// TIA Portal project "智能配药稳定版" (V16)

(* hardware
DEVICE "S7-1200 station_1"  S7-1200 Station
   slot 0: "Rack_0"  S7-1200 Rack  Rack  V1.0
   slot 1: "1.自动供料单元"  CPU 1214C DC/DC/DC  6ES7 214-1AG40-0XB0  V4.4
DEVICE "GSD device_1"  GSD.Device.PN
   slot 0: "机架"  Rack  V1.0
   slot 0: "DEC"  EX-1110  02-01-05  V10.00.00
      slot 0: "TPS Development Toolkit Drivertest"  TPS Development Toolkit Drivertest
      slot 1: "PN-IO"  PN-IO
         slot 1: "Port 1 - RJ45"  Port 1 - RJ45
         slot 2: "Port 2 - RJ45"  Port 2 - RJ45
   slot 1: "EX_210H_1"  EX_210H  1.0
      slot 0: "EX_210H"  EX_210H
   slot 2: "EX_2108_1"  EX_2108  1.0
      slot 0: "EX_2108"  EX_2108
   slot 3: "EX_3208_1"  EX_3208  1.0
      slot 0: "EX_3208"  EX_3208
DEVICE "1.自动供料单元_HMI"  KTP700 Basic PN
   slot 0: "2.自动供料单元_HMI"  KTP700 Basic PN  6AV2 123-2GB03-0AX0  16.0.0.0
   slot 1: "HMI_RT_1"  KTP700 Basic PN  6AV2 123-2GB03-0AX0  16.0.0.0
   slot 5: "2.自动供料单元_HMI.IE_CP_1"  PROFINET Interface  16.0.0.0
      slot 1: "PROFINET Interface_1"  PROFINET Interface
         slot 1: "Port_1"  Port
DEVICE "GSD device_2"  GSD.Device.PN
   slot 0: "机架"  Rack  V1.0
   slot 0: "SINAMICS-V90-PN"  SINAMICS V90 PN V1.0  6SL3 210-5Fxxx-xxFx  V1.00
      slot 0: "SINAMICS V90 PN V1.0"  SINAMICS V90 PN V1.0
      slot 1: "PN-IO"  PN-IO
         slot 1: "端口1"  Port 1
         slot 2: "端口2"  Port 2
      slot 1: "驱动_1"  DRIVE OBJECT
         slot 0: "模块访问点"  Module Access Point
         slot 1: "没有 PROFIsafe"  without PROFIsafe
   slot 2: "标准报文3, PZD-5/9"  Standard telegram 3, PZD 5/9
DEVICE "S7-1200 station_2"  S7-1200 Station
   slot 0: "Rack_0"  S7-1200 Rack  Rack  V1.0
   slot 1: "2.智能分拣单元"  CPU 1214C DC/DC/DC  6ES7 214-1AG40-0XB0  V4.4
DEVICE "2.智能分拣单元_HMI"  KTP700 Basic PN
   slot 0: "HMI_1"  KTP700 Basic PN  6AV2 123-2GB03-0AX0  16.0.0.0
   slot 1: "HMI_RT_2"  KTP700 Basic PN  6AV2 123-2GB03-0AX0  16.0.0.0
   slot 5: "HMI_1.IE_CP_1"  PROFINET Interface  16.0.0.0
      slot 1: "PROFINET Interface_1"  PROFINET Interface
         slot 1: "Port_1"  Port
DEVICE "S7-1200 station_3"  S7-1200 Station
   slot 0: "Rack_0"  S7-1200 Rack  Rack  V1.0
   slot 1: "3.智能仓储单元"  CPU 1214C DC/DC/DC  6ES7 214-1AG40-0XB0  V4.4
   slot 2: "SM 1278_1"  4SI IO link  6ES7 278-4BD32-0XB0  V2.1
   slot 3: "CB 1241 (RS485)"  CB 1241 (RS485)  6ES7 241-1CH30-1XB0  V1.0
   slot 101: "CM 1243-5"  CM 1243-5  6GK7 243-5DX30-0XE0  V1.3
DEVICE "3.智能仓储单元_HMI"  KTP700 Basic PN
   slot 0: "3.智能仓储单元_HMI"  KTP700 Basic PN  6AV2 123-2GB03-0AX0  16.0.0.0
   slot 1: "HMI_RT_3"  KTP700 Basic PN  6AV2 123-2GB03-0AX0  16.0.0.0
   slot 5: "3.智能仓储单元_HMI.IE_CP_1"  PROFINET Interface  16.0.0.0
      slot 1: "PROFINET Interface_1"  PROFINET Interface
         slot 1: "Port_1"  Port
DEVICE "GSD device_3"  GSD.Device.PN
   slot 0: "机架"  Rack  V1.0
   slot 0: "DEC_1"  EX-1110  02-01-05  V10.00.00
      slot 0: "TPS Development Toolkit Drivertest"  TPS Development Toolkit Drivertest
      slot 1: "PN-IO"  PN-IO
         slot 1: "Port 1 - RJ45"  Port 1 - RJ45
         slot 2: "Port 2 - RJ45"  Port 2 - RJ45
   slot 1: "EX_210H_1"  EX_210H  1.0
      slot 0: "EX_210H"  EX_210H
   slot 2: "EX_3208_1"  EX_3208  1.0
      slot 0: "EX_3208"  EX_3208
DEVICE "GSD device_4"  GSD.Device.PN
   slot 0: "机架"  Rack  V1.0
   slot 0: "SINAMICS-V90-PN_1"  SINAMICS V90 PN V1.0  6SL3 210-5Fxxx-xxFx  V1.00
      slot 0: "SINAMICS V90 PN V1.0"  SINAMICS V90 PN V1.0
      slot 1: "PN-IO"  PN-IO
         slot 1: "端口1"  Port 1
         slot 2: "端口2"  Port 2
      slot 1: "驱动_1"  DRIVE OBJECT
         slot 0: "模块访问点"  Module Access Point
         slot 1: "没有 PROFIsafe"  without PROFIsafe
   slot 2: "标准报文3, PZD-5/9"  Standard telegram 3, PZD 5/9
DEVICE "GSD device_5"  GSD.Device.PN
   slot 0: "机架"  Rack  V1.0
   slot 0: "SINAMICS-V90-PN_2"  SINAMICS V90 PN V1.0  6SL3 210-5Fxxx-xxFx  V1.00
      slot 0: "SINAMICS V90 PN V1.0"  SINAMICS V90 PN V1.0
      slot 1: "PN-IO"  PN-IO
         slot 1: "端口1"  Port 1
         slot 2: "端口2"  Port 2
      slot 1: "驱动_1"  DRIVE OBJECT
         slot 0: "模块访问点"  Module Access Point
         slot 1: "没有 PROFIsafe"  without PROFIsafe
   slot 2: "标准报文3, PZD-5/9"  Standard telegram 3, PZD 5/9
DEVICE "GSD device_6"  GSD.Device
   slot 0: "机架_0"  Rail
   slot 0: "Slave_1"  DP-Slave_1  Z1.0
DEVICE "GSD device_7"  GSD.Device.PN
   slot 0: "机架"  Rack  V1.0
   slot 0: "DEC_2"  EX-1110  02-01-05  V10.00.00
      slot 0: "TPS Development Toolkit Drivertest"  TPS Development Toolkit Drivertest
      slot 1: "PN-IO"  PN-IO
         slot 1: "Port 1 - RJ45"  Port 1 - RJ45
         slot 2: "Port 2 - RJ45"  Port 2 - RJ45
   slot 1: "EX_210H_1"  EX_210H  1.0
      slot 0: "EX_210H"  EX_210H
   slot 2: "EX_210H_2"  EX_210H  1.0
      slot 0: "EX_210H"  EX_210H
   slot 3: "EX_3208_1"  EX_3208  1.0
      slot 0: "EX_3208"  EX_3208
   slot 4: "EX_3208_2"  EX_3208  1.0
      slot 0: "EX_3208"  EX_3208
DEVICE "S71500/ET200MP station_1"  S7-1500 station
   slot 0: "导轨_0"  Rack  6ES7 590-1***0-0AA0
   slot 1: "0.数据管理单元"  CPU 1511-1 PN  6ES7 511-1AK02-0AB0  V2.8
      slot 3: "CPU 显示_1"  6ES7591-1AA00-0AA0
      slot 32768: "PROFINET 接口_1"  X1
         slot 32769: "端口_1"  X1 P1
         slot 32770: "端口_2"  X1 P2
      slot 34817: "Virtual CP interface port_1"  Virtual CP interface port  Virtual CP interface port
   slot 2: "DI 16x24VDC / DQ 16x24VDC/0.5A BA_1"  DI 16x24VDC/DQ 16x24VDC/0.5A BA  6ES7 523-1BL00-0AA0  V1.1
DEVICE "GSD device_8"  GSD.Device.PN
   slot 0: "机架"  Rack  V1.0
   slot 0: "SG-GATEWAY"  Master(h750)  SG-PNMB-MS2.0  SW2.0.0
      slot 0: "Master(h750)"  Master(h750)
      slot 1: "X1"  X1
         slot 1: "X1 P1"  X1 P1
         slot 2: "X1 P2"  X1 P2
      slot 1: "Control and Status_1"  Control and Status
         slot 0: "Control and Status"  Control and Status
   slot 2: "03H Read 17 Regs_1"  03H Read 17 Regs
      slot 0: "03H Read 17 Regs"  03H Read 17 Regs
   slot 3: "03H Read 2 Regs_1"  03H Read 2 Regs
      slot 0: "03H Read 2 Regs"  03H Read 2 Regs
   slot 4: "10H Write 1 Reg_1"  10H Write 1 Reg
      slot 0: "10H Write 1 Reg"  10H Write 1 Reg
   slot 5: "03H Read 2 Regs_2"  03H Read 2 Regs
      slot 0: "03H Read 2 Regs"  03H Read 2 Regs
   slot 6: "05H ForceSingleCoil_1"  05H ForceSingleCoil
      slot 0: "05H ForceSingleCoil"  05H ForceSingleCoil
   slot 7: "05H ForceSingleCoil_2"  05H ForceSingleCoil
      slot 0: "05H ForceSingleCoil"  05H ForceSingleCoil
   slot 8: "05H ForceSingleCoil_3"  05H ForceSingleCoil
      slot 0: "05H ForceSingleCoil"  05H ForceSingleCoil
   slot 9: "05H ForceSingleCoil_4"  05H ForceSingleCoil
      slot 0: "05H ForceSingleCoil"  05H ForceSingleCoil
DEVICE "0.数据管理单元_HMI"  KTP700 Basic PN
   slot 0: "0.数据管理单元_HMI"  KTP700 Basic PN  6AV2 123-2GB03-0AX0  16.0.0.0
   slot 1: "HMI_RT_4"  KTP700 Basic PN  6AV2 123-2GB03-0AX0  16.0.0.0
   slot 5: "0.数据管理单元_HMI.IE_CP_1"  PROFINET Interface  16.0.0.0
      slot 1: "PROFINET Interface_1"  PROFINET Interface
         slot 1: "Port_1"  Port
*)

// ===== PLC "1.自动供料单元"  CPU 1214C DC/DC/DC =====

VAR_GLOBAL   // PLC tag table "默认变量表"
   "System_Byte" AT %MB501 : Byte;
   "FirstScan" AT %M501.0 : Bool;
   "DiagStatusUpdate" AT %M501.1 : Bool;
   "AlwaysTRUE" AT %M501.2 : Bool;
   "AlwaysFALSE" AT %M501.3 : Bool;
   "Clock_Byte" AT %MB500 : Byte;
   "Clock_10Hz" AT %M500.0 : Bool;
   "Clock_5Hz" AT %M500.1 : Bool;
   "Clock_2.5Hz" AT %M500.2 : Bool;
   "Clock_2Hz" AT %M500.3 : Bool;
   "Clock_1.25Hz" AT %M500.4 : Bool;
   "Clock_1Hz" AT %M500.5 : Bool;
   "Clock_0.625Hz" AT %M500.6 : Bool;
   "Clock_0.5Hz" AT %M500.7 : Bool;
   "数量检测沿1" AT %M10.0 : Bool;
   "数量检测沿2" AT %M10.1 : Bool;
   "数量检测沿3" AT %M10.2 : Bool;
   "Tag_1" AT %M11.0 : Bool;
   "Tag_2" AT %M11.1 : Bool;
   "Tag_3" AT %M11.2 : Bool;
END_VAR

VAR_GLOBAL   // PLC tag table "第一站变量表"
   "[100]伺服左极限" AT %I0.0 : Bool;
   "[101]伺服右极限" AT %I0.1 : Bool;
   "[102]伺服原点" AT %I0.2 : Bool;
   "[103]步进原点" AT %I0.3 : Bool;
   "[104]步进右极限" AT %I0.4 : Bool;
   "[105]启动" AT %I0.5 : Bool;
   "[106]停止" AT %I0.6 : Bool;
   "[107]复位" AT %I0.7 : Bool;
   "[110]急停" AT %I1.0 : Bool;
   "[111]手自动" AT %I1.1 : Bool;
   "[112]料仓有无料盒" AT %I1.2 : Bool;
   "[113]取料位有无料盒" AT %I1.3 : Bool;
   "[114]功能1" AT %I1.4 : Bool;
   "[115]功能2" AT %I1.5 : Bool;
   "[120]A库物料检测" AT %I2.0 : Bool;
   "[121]B库物料检测" AT %I2.1 : Bool;
   "[122]取料位有无料块" AT %I2.2 : Bool;
   "[123]转盘装配到位检测" AT %I2.3 : Bool;
   "[124]推料盒缩回位" AT %I2.4 : Bool;
   "[125]推料盒伸出位" AT %I2.5 : Bool;
   "[126]A推料伸出位" AT %I2.6 : Bool;
   "[127]A推料缩回位" AT %I2.7 : Bool;
   "[130]B推料伸出位" AT %I3.0 : Bool;
   "[131]B推料缩回位" AT %I3.1 : Bool;
   "[132]取料盒下降位" AT %I3.2 : Bool;
   "[133]取料盒上升位" AT %I3.3 : Bool;
   "[134]取料块伸出位" AT %I3.4 : Bool;
   "[135]取料块缩回位" AT %I3.5 : Bool;
   "[136]取料块下降位" AT %I3.6 : Bool;
   "[137]取料块上升位" AT %I3.7 : Bool;
   "[140]检测伸出位" AT %I4.0 : Bool;
   "[141]检测缩回位" AT %I4.1 : Bool;
   "[142]检测下降位" AT %I4.2 : Bool;
   "[143]检测上升位" AT %I4.3 : Bool;
   "[156]安全光栅" AT %I5.6 : Bool;
   "[164]深度检测当前值" AT %IW64 : Int;
   "轴_1_Drive_IN" AT %I68.0 : "PD_TEL3_IN";
   "[300]转盘步进脉冲" AT %Q0.0 : Bool;
   "[301]转盘步进方向" AT %Q0.1 : Bool;
   "[302]黄色指示灯" AT %Q0.2 : Bool;
   "[303]绿色指示灯" AT %Q0.3 : Bool;
   "[304]红色指示灯" AT %Q0.4 : Bool;
   "[305]转盘皮带电机(正转)" AT %Q0.5 : Bool;
   "[306]转盘皮带电机(反转)" AT %Q0.6 : Bool;
   "[307]声光报警" AT %Q0.7 : Bool;
   "[310]检测伸缩气缸" AT %Q1.0 : Bool;
   "[311]检测升降气缸" AT %Q1.1 : Bool;
   "[320]底盒推料气缸" AT %Q2.0 : Bool;
   "[322]B库推料气缸" AT %Q2.2 : Bool;
   "[323]取底盒升降气缸" AT %Q2.3 : Bool;
   "[324]取料块升降气缸" AT %Q2.4 : Bool;
   "[325]取料块伸缩气缸" AT %Q2.5 : Bool;
   "[326]取料盒夹爪" AT %Q2.6 : Bool;
   "[327]取料块吸盘" AT %Q2.7 : Bool;
   "轴_1_Drive_OUT" AT %Q64.0 : "PD_TEL3_OUT";
   "[144]机械手夹紧到位" AT %I4.4 : Bool;
   "[145]机械手松开到位" AT %I4.5 : Bool;
   "[321]A库推料气缸" AT %Q2.1 : Bool;
END_VAR

DATA_BLOCK "状态控制数据"   // DB33
{ S7_Optimized_Access := 'FALSE' }
VERSION : 0.1
   VAR
      在线状态 : Bool;   // PLC已经上电
      忙碌状态 : Bool;   // 一站已经接单
      空闲状态 : Bool;   // 一站准备就绪(没急停，初始化已经完成，光栅没被挡)
      故障状态 : Bool;   // 报警、光栅被挡
   END_VAR
BEGIN
END_DATA_BLOCK

DATA_BLOCK "初始化数据"   // DB34
{ S7_Optimized_Access := 'FALSE' }
VERSION : 0.1
   VAR
      手动模式 : Bool;
      自动模式 : Bool;
      自动运行模式 : Bool;
      急停状态 : Bool;
      安全光栅被挡 : Bool;
      红灯_内部 : Bool;
      黄灯_内部 : Bool;
      绿灯_内部 : Bool;
      初始化步骤 : Int;
      初始化条件 : Bool;
      初始化下降沿 : Bool;
      初始化中 : Bool;
      初始化故障 : Bool;
      初始化完成 : Bool;
      报警等级 : Int;
      报警确认按钮 : Bool;
      气缸报警复位 : Bool;
      底盒推料气缸报警 : Bool;
      A库推料气缸报警 : Bool;
      B库推料气缸报警 : Bool;
      检测伸缩气缸报警 : Bool;
      检测升降气缸报警 : Bool;
      取料块升降气缸报警 : Bool;
      取料块伸缩气缸报警 : Bool;
      取料盒夹爪报警 : Bool;
      气缸报警输出 : Bool;
      轴回零错误 : Bool;
      报警总输出 : Bool;
   END_VAR
BEGIN
END_DATA_BLOCK

// folder: System blocks/Program resources

DATA_BLOCK "吸住料块上升计时"   // DB10
{ S7_Optimized_Access := 'TRUE' }
AUTHOR : Simatic
FAMILY : IEC
NAME : IEC_TMR
VERSION : 1.0
// stored: InstanceOfName IEC_TIMER
"IEC_TIMER"
BEGIN
END_DATA_BLOCK

DATA_BLOCK "IEC_Timer_0_DB_10"   // DB14
{ S7_Optimized_Access := 'TRUE' }
AUTHOR : Simatic
FAMILY : IEC
NAME : IEC_TMR
VERSION : 1.0
// stored: InstanceOfName IEC_TIMER
"IEC_TIMER"
BEGIN
END_DATA_BLOCK

DATA_BLOCK "IEC_Timer_0_DB_5"   // DB16
{ S7_Optimized_Access := 'TRUE' }
AUTHOR : Simatic
FAMILY : IEC
NAME : IEC_TMR
VERSION : 1.0
// stored: InstanceOfName IEC_TIMER
"IEC_TIMER"
BEGIN
END_DATA_BLOCK

DATA_BLOCK "IEC_Timer_0_DB_2"   // DB19
{ S7_Optimized_Access := 'TRUE' }
AUTHOR : Simatic
FAMILY : IEC
NAME : IEC_TMR
VERSION : 1.0
// stored: InstanceOfName IEC_TIMER
"IEC_TIMER"
BEGIN
END_DATA_BLOCK

DATA_BLOCK "IEC_Timer_0_DB_3"   // DB21
{ S7_Optimized_Access := 'TRUE' }
AUTHOR : Simatic
FAMILY : IEC
NAME : IEC_TMR
VERSION : 1.0
// stored: InstanceOfName IEC_TIMER
"IEC_TIMER"
BEGIN
END_DATA_BLOCK

DATA_BLOCK "IEC_Timer_0_DB_7"   // DB23
{ S7_Optimized_Access := 'TRUE' }
AUTHOR : Simatic
FAMILY : IEC
NAME : IEC_TMR
VERSION : 1.0
// stored: InstanceOfName IEC_TIMER
"IEC_TIMER"
BEGIN
END_DATA_BLOCK

DATA_BLOCK "IEC_Timer_0_DB_6"   // DB24
{ S7_Optimized_Access := 'TRUE' }
AUTHOR : Simatic
FAMILY : IEC
NAME : IEC_TMR
VERSION : 1.0
// stored: InstanceOfName IEC_TIMER
"IEC_TIMER"
BEGIN
END_DATA_BLOCK

DATA_BLOCK "IEC_Timer_0_DB_8"   // DB25
{ S7_Optimized_Access := 'TRUE' }
AUTHOR : Simatic
FAMILY : IEC
NAME : IEC_TMR
VERSION : 1.0
// stored: InstanceOfName IEC_TIMER
"IEC_TIMER"
BEGIN
END_DATA_BLOCK

DATA_BLOCK "IEC_Timer_0_DB_9"   // DB26
{ S7_Optimized_Access := 'TRUE' }
AUTHOR : Simatic
FAMILY : IEC
NAME : IEC_TMR
VERSION : 1.0
// stored: InstanceOfName IEC_TIMER
"IEC_TIMER"
BEGIN
END_DATA_BLOCK

DATA_BLOCK "IEC_Timer_0_DB_11"   // DB27
{ S7_Optimized_Access := 'TRUE' }
AUTHOR : Simatic
FAMILY : IEC
NAME : IEC_TMR
VERSION : 1.0
// stored: InstanceOfName IEC_TIMER
"IEC_TIMER"
BEGIN
END_DATA_BLOCK

DATA_BLOCK "IEC_Timer_0_DB_12"   // DB28
{ S7_Optimized_Access := 'TRUE' }
AUTHOR : Simatic
FAMILY : IEC
NAME : IEC_TMR
VERSION : 1.0
// stored: InstanceOfName IEC_TIMER
"IEC_TIMER"
BEGIN
END_DATA_BLOCK

DATA_BLOCK "IEC_Timer_0_DB_13"   // DB29
{ S7_Optimized_Access := 'TRUE' }
AUTHOR : Simatic
FAMILY : IEC
NAME : IEC_TMR
VERSION : 1.0
// stored: InstanceOfName IEC_TIMER
"IEC_TIMER"
BEGIN
END_DATA_BLOCK

DATA_BLOCK "IEC_Timer_0_DB_14"   // DB30
{ S7_Optimized_Access := 'TRUE' }
AUTHOR : Simatic
FAMILY : IEC
NAME : IEC_TMR
VERSION : 1.0
// stored: InstanceOfName IEC_TIMER
"IEC_TIMER"
BEGIN
END_DATA_BLOCK

DATA_BLOCK "IEC_Timer_0_DB_15"   // DB31
{ S7_Optimized_Access := 'TRUE' }
AUTHOR : Simatic
FAMILY : IEC
NAME : IEC_TMR
VERSION : 1.0
// stored: InstanceOfName IEC_TIMER
"IEC_TIMER"
BEGIN
END_DATA_BLOCK

DATA_BLOCK "IEC_Timer_0_DB_4"   // DB32
{ S7_Optimized_Access := 'TRUE' }
AUTHOR : Simatic
FAMILY : IEC
NAME : IEC_TMR
VERSION : 1.0
// stored: InstanceOfName IEC_TIMER
"IEC_TIMER"
BEGIN
END_DATA_BLOCK

DATA_BLOCK "IEC_Timer_0_DB_23"   // DB35
{ S7_Optimized_Access := 'TRUE' }
AUTHOR : Simatic
FAMILY : IEC
NAME : IEC_TMR
VERSION : 1.0
// stored: InstanceOfName IEC_TIMER
"IEC_TIMER"
BEGIN
END_DATA_BLOCK

DATA_BLOCK "_1.自动供料单元_Receive_DB"   // DB38
{ S7_Optimized_Access := 'TRUE' }
AUTHOR : SIMATIC
FAMILY : MC7Plus
NAME : TC_IP_v4
VERSION : 1.0
// stored: InstanceOfName TCON_IP_v4
"TCON_IP_v4"
BEGIN
   ID := 105;
   InterfaceId := 64;
   LocalPort := 8899;
   RemotePort := 8899;
   RemoteAddress.ADDR[1] := 192;
   RemoteAddress.ADDR[2] := 168;
   RemoteAddress.ADDR[3] := 40;
   RemoteAddress.ADDR[4] := 100;
END_DATA_BLOCK

DATA_BLOCK "IEC_Timer_0_DB_24"   // DB39
{ S7_Optimized_Access := 'TRUE' }
AUTHOR : Simatic
FAMILY : IEC
NAME : IEC_TMR
VERSION : 1.0
// stored: InstanceOfName IEC_TIMER
"IEC_TIMER"
BEGIN
END_DATA_BLOCK

DATA_BLOCK "IEC_Timer_0_DB_16"   // DB40
{ S7_Optimized_Access := 'TRUE' }
AUTHOR : Simatic
FAMILY : IEC
NAME : IEC_TMR
VERSION : 1.0
// stored: InstanceOfName IEC_TIMER
"IEC_TIMER"
BEGIN
END_DATA_BLOCK

DATA_BLOCK "IEC_Timer_0_DB_17"   // DB41
{ S7_Optimized_Access := 'TRUE' }
AUTHOR : Simatic
FAMILY : IEC
NAME : IEC_TMR
VERSION : 1.0
// stored: InstanceOfName IEC_TIMER
"IEC_TIMER"
BEGIN
END_DATA_BLOCK

DATA_BLOCK "IEC_Timer_0_DB_18"   // DB42
{ S7_Optimized_Access := 'TRUE' }
AUTHOR : Simatic
FAMILY : IEC
NAME : IEC_TMR
VERSION : 1.0
// stored: InstanceOfName IEC_TIMER
"IEC_TIMER"
BEGIN
END_DATA_BLOCK

DATA_BLOCK "IEC_Timer_0_DB_19"   // DB43
{ S7_Optimized_Access := 'TRUE' }
AUTHOR : Simatic
FAMILY : IEC
NAME : IEC_TMR
VERSION : 1.0
// stored: InstanceOfName IEC_TIMER
"IEC_TIMER"
BEGIN
END_DATA_BLOCK

DATA_BLOCK "IEC_Timer_0_DB_20"   // DB44
{ S7_Optimized_Access := 'TRUE' }
AUTHOR : Simatic
FAMILY : IEC
NAME : IEC_TMR
VERSION : 1.0
// stored: InstanceOfName IEC_TIMER
"IEC_TIMER"
BEGIN
END_DATA_BLOCK

DATA_BLOCK "IEC_Timer_0_DB_21"   // DB45
{ S7_Optimized_Access := 'TRUE' }
AUTHOR : Simatic
FAMILY : IEC
NAME : IEC_TMR
VERSION : 1.0
// stored: InstanceOfName IEC_TIMER
"IEC_TIMER"
BEGIN
END_DATA_BLOCK

DATA_BLOCK "IEC_Timer_0_DB_22"   // DB46
{ S7_Optimized_Access := 'TRUE' }
AUTHOR : Simatic
FAMILY : IEC
NAME : IEC_TMR
VERSION : 1.0
// stored: InstanceOfName IEC_TIMER
"IEC_TIMER"
BEGIN
END_DATA_BLOCK

// folder: 手动模式

DATA_BLOCK "手动模式数据"   // DB12
{ S7_Optimized_Access := 'FALSE' }
VERSION : 0.1
   VAR
      S10推料盒步骤 : Real;
      S20推料块步骤 : Real;
      S30放料块步骤 : Real;
      S40送料盒步骤 : Real;
      手动总步骤 : Real;
      料块仓选择 : Int := 1;
      沿1 : Bool;
      沿2 : Bool;
      沿3 : Bool;
      沿4 : Bool;
   END_VAR
BEGIN
END_DATA_BLOCK

// folder: 自动模式

DATA_BLOCK "自动模式数据"   // DB22
{ S7_Optimized_Access := 'FALSE' }
VERSION : 0.1
   VAR
      Z10步骤 : Real;
      Z20步骤 : Real;
      Z30步骤 : Real;
      Z40步骤 : Real;
      Z50步骤 : Real;
      自动模式总步骤 : Real;
      推料盒数 : Bool;
      开始信号 : Bool;
      ab物料选择 : Int;
      料盒使用数 : Int;
      a料使用数 : Int;
      b料使用数 : Int;
      当前深度检测_1 : Real;   // 模数转换
      当前深度检测_2 : Real;   // 模数转换
      当前深度检测 : Real;
      深度保存 : Array[0..1] of Real;
      扫码器接受数据 : String[16];
      扫码器扫码数值 : Int;
      扫码器扫码成功 : Bool;
   END_VAR
BEGIN
END_DATA_BLOCK

// folder: 运动控制

DATA_BLOCK "运动控制数据块"   // DB1
{ S7_Optimized_Access := 'FALSE' }
VERSION : 0.1
   VAR
      转盘目标角度 : Real;
      转盘目标速度 : Real;
      转盘实际角度 : Real;
      转盘实际速度 : Real;
      转盘步进使能 : Bool;
      转盘步进使能状态 : Bool;
      转盘使能错误 : Bool;
      转盘复位按钮 : Bool;
      转盘复位完成 : Bool;
      转盘复位错误 : Bool;
      转盘回原点按钮 : Bool;
      转盘回原点完成 : Bool;
      转盘回原点错误 : Bool;
      转盘绝对定位按钮 : Bool;
      转盘绝对定位完成 : Bool;
      转盘绝对定位错误 : Bool;
      机械手目标位置 : Real;
      机械手目标速度 : Real;
      机械手实际位置 : Real;
      机械手实际速度 : Real;
      机械手伺服使能 : Bool;
      机械手伺服使能状态 : Bool;
      机械手使能错误 : Bool;
      机械手复位按钮 : Bool;
      机械手复位完成 : Bool;
      机械手复位错误 : Bool;
      机械手回原点按钮 : Bool;
      机械手回原点完成 : Bool;
      机械手回原点错误 : Bool;
      机械手绝对定位按钮 : Bool;
      机械手绝对定位完成 : Bool;
      机械手绝对定位错误 : Bool;
      机械手左移点动 : Bool;
      机械手右移点动 : Bool;
      轴初始化按钮 : Bool;
      轴初始化完成 : Bool;
      轴初始化步骤 : Int;
      轴初始化错误 : Bool;
      转盘轴错误输出 : Bool;
      机械手轴错误输出 : Bool;
   END_VAR
BEGIN
END_DATA_BLOCK

// folder: 通讯数据

DATA_BLOCK "虚实联动信号"   // DB109
{ S7_Optimized_Access := 'FALSE' }
VERSION : 0.1
   VAR
      底盒推料气缸 : Bool;
      皮带正转 : Bool;
      皮带反转 : Bool;
      A库推料气缸 : Bool;
      B库推料气缸 : Bool;
      取底盒升降气缸 : Bool;
      取料盒夹爪 : Bool;
      一站机械手位置 : Real;
      一站机械手速度 : Real;
      转盘角度 : Real;
      转盘速度 : Real;
      取料块吸盘 : Bool;
      取料块升降气缸 : Bool;
      取料块伸缩气缸 : Bool;
      检测伸缩气缸 : Bool;
      检测升降气缸 : Bool;
   END_VAR
BEGIN
END_DATA_BLOCK

DATA_BLOCK "一站数据"   // DB111
{ S7_Optimized_Access := 'FALSE' }
VERSION : 0.1
   VAR
      一站完成 : Bool;
      复位完成 : Bool;
      一站就绪 : Bool;
      一站忙碌 : Bool;
      一站请求二站接收 : Bool;
      一站可接单 : Bool;
      数据7 : Bool;
      数据8 : Bool;
      数据9 : Bool;
      数据10 : Bool;
      数据11 : Bool;
      数据12 : Bool;
      数据13 : Bool;
      数据14 : Bool;
   END_VAR
BEGIN
END_DATA_BLOCK

DATA_BLOCK "二站数据"   // DB112
{ S7_Optimized_Access := 'FALSE' }
VERSION : 0.1
   VAR
      二站完成 : Bool;
      二站已接收 : Bool;
      复位完成 : Bool;
      空闲状态 : Bool;
      电机正转 : Bool;
      二站忙碌 : Bool;
      二站请求三站接收 : Bool;
      二站可接收 : Bool;
      数据17 : Bool;
      数据18 : Bool;
      数据19 : Bool;
      数据20 : Bool;
      数据21 : Bool;
   END_VAR
BEGIN
END_DATA_BLOCK

DATA_BLOCK "AI通讯数据"   // DB116
{ S7_Optimized_Access := 'FALSE' }
VERSION : 0.1
   VAR
      一站上料到位 : Bool;
      一站压装到位 : Bool;
   END_VAR
BEGIN
END_DATA_BLOCK

DATA_BLOCK "一站MES读取数据"   // DB120
{ S7_Optimized_Access := 'FALSE' }
VERSION : 0.1
   VAR
      一站数据 : Struct
         在线状态 : Int;
         运行模式 : Int;   // 0 手动 / 1 自动待机 / 2 自动运行
         忙碌状态 : Int;   // 0 空闲 / 1 忙碌
         故障状态 : Int;   // 0 = 无故障
         当前订单ID : Int;   // 当前处理的订单
         当前步骤 : Real;
         心跳值 : Int;
         一站完成 : Bool;
         订单完成一站复位 : Bool;
         保留_1 : Bool;
         保留_2 : Bool;
         保留_3 : Bool;
         保留_4 : Bool;
         保留_5 : Bool;
         保留_6 : Bool;
         扫码条码数据 : Int;
         转盘当前角度 : Real;
         机械手当前位置 : Real;
         深度检测值 : Real;
         料盒使用数 : Int;
         A料使用数 : Int;
         B料使用数 : Int;
         一站保留数据 : Array[0..9] of Int;
      END_STRUCT;
      订单数据 : Struct
         订单id : Int;
         ab物料 : Int;   // 1A，2B，3不需要
         小钢珠数量 : Int;
         大钢珠数量 : Int;
         存储仓位 : Int;
         当前订单完成 : Bool;
         开始信号 : Int;
         复位信号 : Int;
         订单保留数据 : Array[0..4] of Int;
      END_STRUCT;
   END_VAR
BEGIN
END_DATA_BLOCK

// folder: (top level)

DATA_BLOCK "机械手"   // DB2, Motion_DB
{ S7_Optimized_Access := 'TRUE' }
AUTHOR : SIMATIC
FAMILY : BasicMC
NAME : TO_PosAx
VERSION : 7.0
// stored: InstanceOfName TO_PositioningAxis
"TO_PositioningAxis"
BEGIN
   // Axis.Encoder.TelegramAddressOutCU = %Q64.0
   // Axis.Encoder.TelegramAddressInCU = %I68.0
   // Axis.Encoder.DoNameCU = SINAMICS-V90-PN.驱动_1_编码器1
   // Axis.Drive.TelegramAddressOutCU = %Q64.0
   // Axis.Drive.TelegramAddressInCU = %I68.0
   // Axis.Drive.TelegramType = 2
   // Axis.Drive.DoNameCU = SINAMICS-V90-PN.驱动_1
   // Axis.HomingReferencePointSwitch_AddressCU = %I0.2
   // Axis.PositionLimitsMax_AddressCU = %I0.0
   // Axis.PositionLimitsMin_AddressCU = %I0.1
   // Axis.LengthUnitNormalized.Distance = 1013
   // Axis.Encoder.SelectedHscIndexCU = -1
   // Axis.Encoder.DbTypeCU = Classic
   // Axis.Drive.DbTypeCU = Classic
END_DATA_BLOCK

DATA_BLOCK "转盘"   // DB3, Motion_DB
{ S7_Optimized_Access := 'TRUE' }
AUTHOR : SIMATIC
FAMILY : BasicMC
NAME : TO_PosAx
VERSION : 7.0
// stored: InstanceOfName TO_PositioningAxis
"TO_PositioningAxis"
BEGIN
   // Axis.HomingReferencePointSwitch_AddressCU = %I0.3
   // Axis.LengthUnitNormalized.Distance = 1005
   // Axis.LengthUnit.LastDistance = 1005
   // Axis.PositionLimitsMax_AddressCU = %I0.4
   // Axis.PositionLimitsMin_AddressCU = %I0.0
   // Axis.DirectionOutputEnabledCU = TRUE
   // Axis.OnlinePtoModeCU = 16#0000_0002
   // Axis.SelectedChannel2EnumCU = %Q0.1
   // Axis.SelectedChannel1EnumCU = %Q0.0
   // Pulse.MinDeltaDeltaFrequencyCU = 0.004
   // Pulse.MaxDeltaDeltaFrequencyCU = 1.0E+10
   // Pulse.MinDeltaFrequencyCU = 0.005
   // Pulse.MaxDeltaFrequencyCU = 9.5E+9
   // Pulse.MinFrequencyCU = 1.0
   // Pulse.MaxFrequencyCU = 100000.0
   // Pulse.OutputSourceCU = 16#0000_0000
   // Axis.SelectPTO = 0
END_DATA_BLOCK

FUNCTION "1.报警程序" : Void   // FC10, LAD
{ S7_Optimized_Access := 'TRUE' }
VERSION : 0.1
BEGIN

REGION Network 1: 气缸报警——————底盒推料气缸
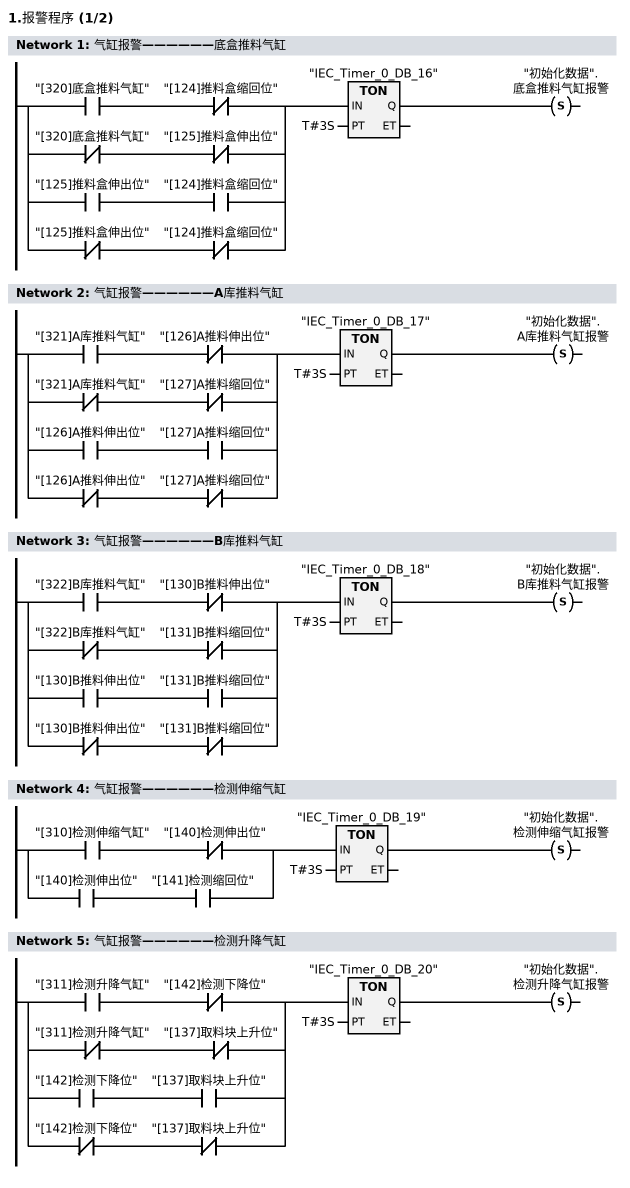
   "IEC_Timer_0_DB_16".TON(IN := ("[320]底盒推料气缸" AND NOT "[124]推料盒缩回位") OR (NOT "[320]底盒推料气缸" AND NOT "[125]推料盒伸出位") OR ("[125]推料盒伸出位" AND "[124]推料盒缩回位") OR (NOT "[125]推料盒伸出位" AND NOT "[124]推料盒缩回位"),
                           PT := T#3S);
   IF "IEC_Timer_0_DB_16".Q THEN "初始化数据".底盒推料气缸报警 := TRUE; END_IF;
END_REGION

REGION Network 2: 气缸报警——————A库推料气缸
   "IEC_Timer_0_DB_17".TON(IN := ("[321]A库推料气缸" AND NOT "[126]A推料伸出位") OR (NOT "[321]A库推料气缸" AND NOT "[127]A推料缩回位") OR ("[126]A推料伸出位" AND "[127]A推料缩回位") OR (NOT "[126]A推料伸出位" AND NOT "[127]A推料缩回位"),
                           PT := T#3S);
   IF "IEC_Timer_0_DB_17".Q THEN "初始化数据".A库推料气缸报警 := TRUE; END_IF;
END_REGION

REGION Network 3: 气缸报警——————B库推料气缸
   "IEC_Timer_0_DB_18".TON(IN := ("[322]B库推料气缸" AND NOT "[130]B推料伸出位") OR (NOT "[322]B库推料气缸" AND NOT "[131]B推料缩回位") OR ("[130]B推料伸出位" AND "[131]B推料缩回位") OR (NOT "[130]B推料伸出位" AND NOT "[131]B推料缩回位"),
                           PT := T#3S);
   IF "IEC_Timer_0_DB_18".Q THEN "初始化数据".B库推料气缸报警 := TRUE; END_IF;
END_REGION

REGION Network 4: 气缸报警——————检测伸缩气缸
   "IEC_Timer_0_DB_19".TON(IN := ("[310]检测伸缩气缸" AND NOT "[140]检测伸出位") OR ("[140]检测伸出位" AND "[141]检测缩回位"),
                           PT := T#3S);
   IF "IEC_Timer_0_DB_19".Q THEN "初始化数据".检测伸缩气缸报警 := TRUE; END_IF;
END_REGION

REGION Network 5: 气缸报警——————检测升降气缸
   "IEC_Timer_0_DB_20".TON(IN := ("[311]检测升降气缸" AND NOT "[142]检测下降位") OR (NOT "[311]检测升降气缸" AND NOT "[137]取料块上升位") OR ("[142]检测下降位" AND "[137]取料块上升位") OR (NOT "[142]检测下降位" AND NOT "[137]取料块上升位"),
                           PT := T#3S);
   IF "IEC_Timer_0_DB_20".Q THEN "初始化数据".检测升降气缸报警 := TRUE; END_IF;
END_REGION

REGION Network 6: 气缸报警——————取料块升降气缸
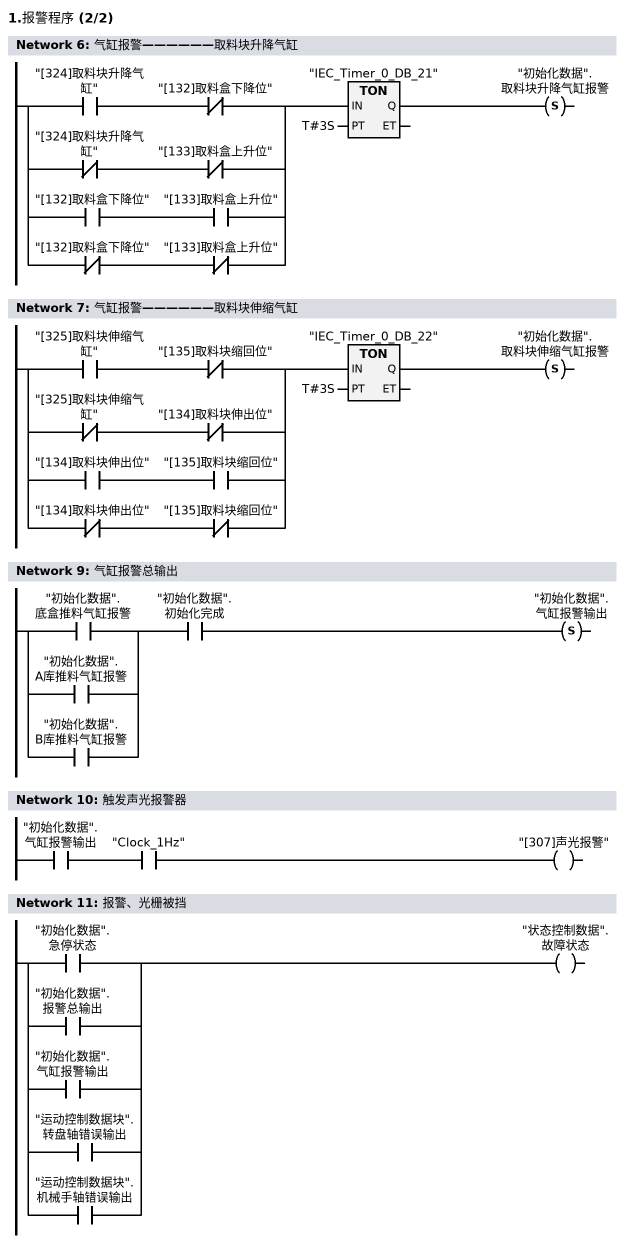
   "IEC_Timer_0_DB_21".TON(IN := ("[324]取料块升降气缸" AND NOT "[132]取料盒下降位") OR (NOT "[324]取料块升降气缸" AND NOT "[133]取料盒上升位") OR ("[132]取料盒下降位" AND "[133]取料盒上升位") OR (NOT "[132]取料盒下降位" AND NOT "[133]取料盒上升位"),
                           PT := T#3S);
   IF "IEC_Timer_0_DB_21".Q THEN "初始化数据".取料块升降气缸报警 := TRUE; END_IF;
END_REGION

REGION Network 7: 气缸报警——————取料块伸缩气缸
   "IEC_Timer_0_DB_22".TON(IN := ("[325]取料块伸缩气缸" AND NOT "[135]取料块缩回位") OR (NOT "[325]取料块伸缩气缸" AND NOT "[134]取料块伸出位") OR ("[134]取料块伸出位" AND "[135]取料块缩回位") OR (NOT "[134]取料块伸出位" AND NOT "[135]取料块缩回位"),
                           PT := T#3S);
   IF "IEC_Timer_0_DB_22".Q THEN "初始化数据".取料块伸缩气缸报警 := TRUE; END_IF;
END_REGION

REGION Network 9: 气缸报警总输出
   RUNG wire#powerrail
      Contact( "初始化数据".底盒推料气缸报警 )
      wire#w1
      Contact( "初始化数据".初始化完成 )
      S_Coil( "初始化数据".气缸报警输出 )
   END_RUNG
   RUNG wire#powerrail
      Contact( "初始化数据".A库推料气缸报警 )
   END_RUNG wire#w1
   RUNG wire#powerrail
      Contact( "初始化数据".B库推料气缸报警 )
   END_RUNG wire#w1
   // the same network as SCL:
   IF ("初始化数据".底盒推料气缸报警 OR "初始化数据".A库推料气缸报警 OR "初始化数据".B库推料气缸报警) AND "初始化数据".初始化完成 THEN
       "初始化数据".气缸报警输出 := TRUE;
   END_IF;
END_REGION

REGION Network 10: 触发声光报警器
   RUNG wire#powerrail
      Contact( "初始化数据".气缸报警输出 )
      Contact( "Clock_1Hz" )
      Coil( "[307]声光报警" )
   END_RUNG
   // the same network as SCL:
   "[307]声光报警" := "初始化数据".气缸报警输出 AND "Clock_1Hz";
END_REGION

REGION Network 11: 报警、光栅被挡
   RUNG wire#powerrail
      Contact( "初始化数据".急停状态 )
      wire#w1
      Coil( "状态控制数据".故障状态 )
   END_RUNG
   RUNG wire#powerrail
      Contact( "初始化数据".报警总输出 )
   END_RUNG wire#w1
   RUNG wire#powerrail
      Contact( "初始化数据".气缸报警输出 )
   END_RUNG wire#w1
   RUNG wire#powerrail
      Contact( "运动控制数据块".转盘轴错误输出 )
   END_RUNG wire#w1
   RUNG wire#powerrail
      Contact( "运动控制数据块".机械手轴错误输出 )
   END_RUNG wire#w1
   // the same network as SCL:
   "状态控制数据".故障状态 := "初始化数据".急停状态 OR "初始化数据".报警总输出 OR "初始化数据".气缸报警输出 OR "运动控制数据块".转盘轴错误输出 OR "运动控制数据块".机械手轴错误输出;
END_REGION
END_FUNCTION

FUNCTION "0.初始化" : Void   // FC13, LAD
{ S7_Optimized_Access := 'TRUE' }
VERSION : 0.1
   VAR_TEMP   // added for the SCL form of the ladder/FBD networks
      _w1 : Bool;
      _w2 : Bool;
   END_VAR
BEGIN

REGION Network 1: 模式切换
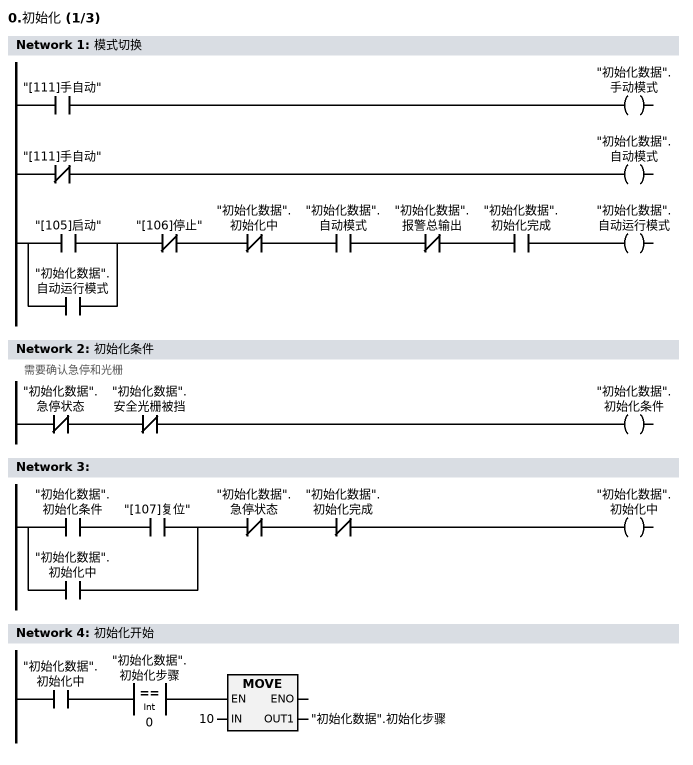
   RUNG wire#powerrail
      Contact( "[111]手自动" )
      Coil( "初始化数据".手动模式 )
   END_RUNG
   RUNG wire#powerrail
      I_Contact( "[111]手自动" )
      Coil( "初始化数据".自动模式 )
   END_RUNG
   RUNG wire#powerrail
      Contact( "[105]启动" )
      wire#w1
      I_Contact( "[106]停止" )
      I_Contact( "初始化数据".初始化中 )
      Contact( "初始化数据".自动模式 )
      I_Contact( "初始化数据".报警总输出 )
      Contact( "初始化数据".初始化完成 )
      Coil( "初始化数据".自动运行模式 )
   END_RUNG
   RUNG wire#powerrail
      Contact( "初始化数据".自动运行模式 )
   END_RUNG wire#w1
   // the same network as SCL:
   "初始化数据".手动模式 := "[111]手自动";
   "初始化数据".自动模式 := NOT "[111]手自动";
   "初始化数据".自动运行模式 := ("[105]启动" OR "初始化数据".自动运行模式) AND NOT "[106]停止" AND NOT "初始化数据".初始化中 AND "初始化数据".自动模式 AND NOT "初始化数据".报警总输出 AND "初始化数据".初始化完成;
END_REGION

REGION Network 2: 初始化条件
   // 需要确认急停和光栅
   RUNG wire#powerrail
      I_Contact( "初始化数据".急停状态 )
      I_Contact( "初始化数据".安全光栅被挡 )
      Coil( "初始化数据".初始化条件 )
   END_RUNG
   // the same network as SCL:
   "初始化数据".初始化条件 := NOT "初始化数据".急停状态 AND NOT "初始化数据".安全光栅被挡;
END_REGION

REGION Network 3
   RUNG wire#powerrail
      Contact( "初始化数据".初始化条件 )
      Contact( "[107]复位" )
      wire#w1
      I_Contact( "初始化数据".急停状态 )
      I_Contact( "初始化数据".初始化完成 )
      Coil( "初始化数据".初始化中 )
   END_RUNG
   RUNG wire#powerrail
      Contact( "初始化数据".初始化中 )
   END_RUNG wire#w1
   // the same network as SCL:
   "初始化数据".初始化中 := (("初始化数据".初始化条件 AND "[107]复位") OR "初始化数据".初始化中) AND NOT "初始化数据".急停状态 AND NOT "初始化数据".初始化完成;
END_REGION

REGION Network 4: 初始化开始
   RUNG wire#powerrail
      Contact( "初始化数据".初始化中 )
      { S7_Templates := "SrcType := Int" } EQ_Contact(in1 := "初始化数据".初始化步骤, in2 := 0)
      Move(in := 10, out1 => "初始化数据".初始化步骤)
   END_RUNG
   // the same network as SCL:
   IF "初始化数据".初始化中 AND ("初始化数据".初始化步骤 = 0) THEN "初始化数据".初始化步骤 := 10; END_IF;
END_REGION

REGION Network 5: 数据初始化
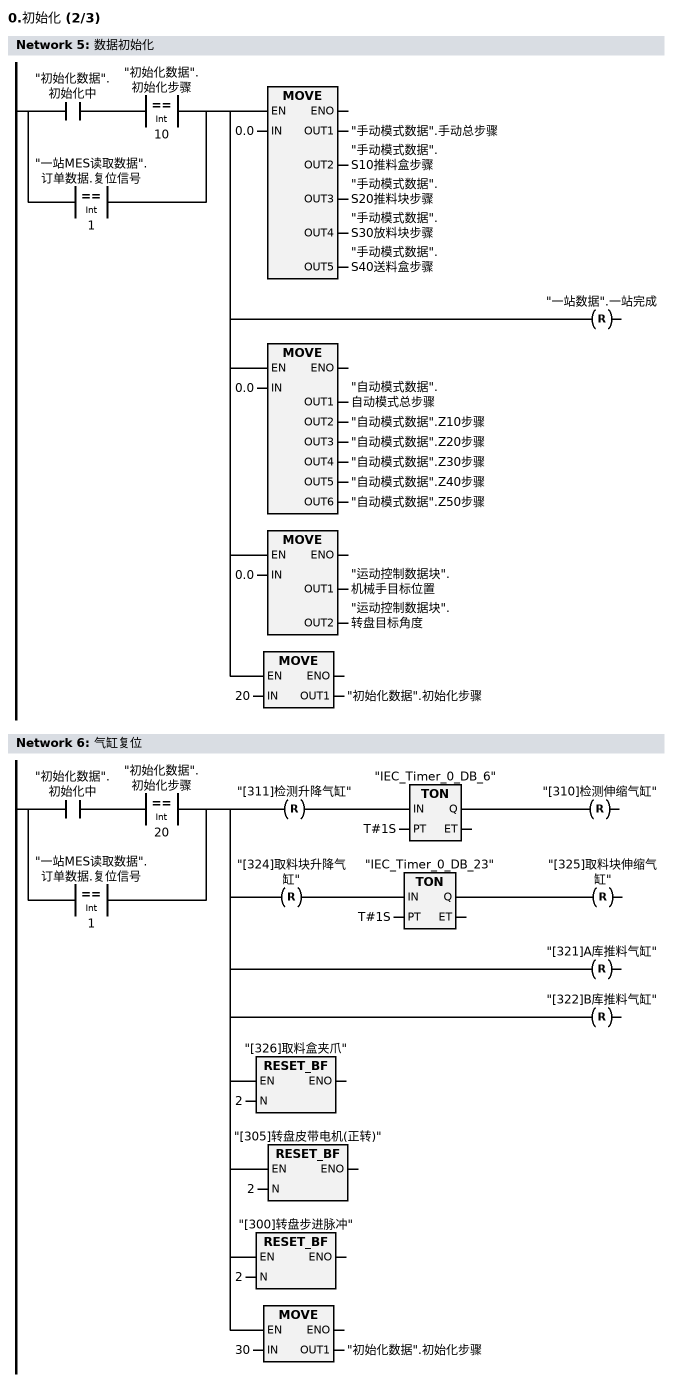
   RUNG wire#powerrail
      Contact( "初始化数据".初始化中 )
      { S7_Templates := "SrcType := Int" } EQ_Contact(in1 := "初始化数据".初始化步骤, in2 := 10)
      wire#w1
      Move(in := 0.0, out1 => "手动模式数据".手动总步骤, out2 => "手动模式数据".S10推料盒步骤, out3 => "手动模式数据".S20推料块步骤, out4 => "手动模式数据".S30放料块步骤, out5 => "手动模式数据".S40送料盒步骤)
   END_RUNG
   RUNG wire#powerrail
      { S7_Templates := "SrcType := Int" } EQ_Contact(in1 := "一站MES读取数据".订单数据.复位信号, in2 := 1)
   END_RUNG wire#w1
   RUNG wire#w1
      R_Coil( "一站数据".一站完成 )
   END_RUNG
   RUNG wire#w1
      Move(in := 0.0, out1 => "自动模式数据".自动模式总步骤, out2 => "自动模式数据".Z10步骤, out3 => "自动模式数据".Z20步骤, out4 => "自动模式数据".Z30步骤, out5 => "自动模式数据".Z40步骤, out6 => "自动模式数据".Z50步骤)
   END_RUNG
   RUNG wire#w1
      Move(in := 0.0, out1 => "运动控制数据块".机械手目标位置, out2 => "运动控制数据块".转盘目标角度)
   END_RUNG
   RUNG wire#w1
      Move(in := 20, out1 => "初始化数据".初始化步骤)
   END_RUNG
   // the same network as SCL:
   IF ("初始化数据".初始化中 AND ("初始化数据".初始化步骤 = 10)) OR ("一站MES读取数据".订单数据.复位信号 = 1) THEN
       "手动模式数据".手动总步骤 := 0.0;
       "手动模式数据".S10推料盒步骤 := 0.0;
       "手动模式数据".S20推料块步骤 := 0.0;
       "手动模式数据".S30放料块步骤 := 0.0;
       "手动模式数据".S40送料盒步骤 := 0.0;
       "一站数据".一站完成 := FALSE;
       "自动模式数据".自动模式总步骤 := 0.0;
       "自动模式数据".Z10步骤 := 0.0;
       "自动模式数据".Z20步骤 := 0.0;
       "自动模式数据".Z30步骤 := 0.0;
       "自动模式数据".Z40步骤 := 0.0;
       "自动模式数据".Z50步骤 := 0.0;
       "运动控制数据块".机械手目标位置 := 0.0;
       "运动控制数据块".转盘目标角度 := 0.0;
       "初始化数据".初始化步骤 := 20;
   END_IF;
END_REGION

REGION Network 6: 气缸复位
   // no SCL statement known for RBitfield: written as a call
   #_w1 := ("初始化数据".初始化中 AND ("初始化数据".初始化步骤 = 20)) OR ("一站MES读取数据".订单数据.复位信号 = 1);
   IF #_w1 THEN "[311]检测升降气缸" := FALSE; END_IF;
   "IEC_Timer_0_DB_6".TON(IN := #_w1, PT := T#1S);
   IF "IEC_Timer_0_DB_6".Q THEN "[310]检测伸缩气缸" := FALSE; END_IF;
   IF #_w1 THEN "[324]取料块升降气缸" := FALSE; END_IF;
   "IEC_Timer_0_DB_23".TON(IN := #_w1, PT := T#1S);
   IF "IEC_Timer_0_DB_23".Q THEN "[325]取料块伸缩气缸" := FALSE; END_IF;
   IF #_w1 THEN
       "[321]A库推料气缸" := FALSE;
       "[322]B库推料气缸" := FALSE;
       RESET_BF(operand := "[326]取料盒夹爪", n := 2);
       RESET_BF(operand := "[305]转盘皮带电机(正转)", n := 2);
       RESET_BF(operand := "[300]转盘步进脉冲", n := 2);
       "初始化数据".初始化步骤 := 30;
   END_IF;
END_REGION

REGION Network 7: 轴复位
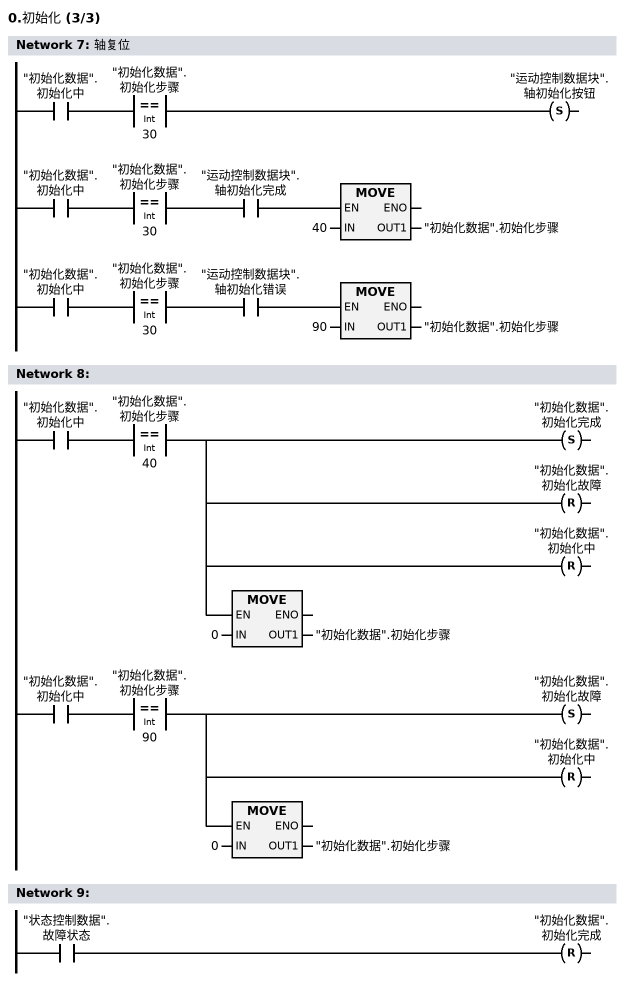
   RUNG wire#powerrail
      Contact( "初始化数据".初始化中 )
      { S7_Templates := "SrcType := Int" } EQ_Contact(in1 := "初始化数据".初始化步骤, in2 := 30)
      S_Coil( "运动控制数据块".轴初始化按钮 )
   END_RUNG
   RUNG wire#powerrail
      Contact( "初始化数据".初始化中 )
      { S7_Templates := "SrcType := Int" } EQ_Contact(in1 := "初始化数据".初始化步骤, in2 := 30)
      Contact( "运动控制数据块".轴初始化完成 )
      Move(in := 40, out1 => "初始化数据".初始化步骤)
   END_RUNG
   RUNG wire#powerrail
      Contact( "初始化数据".初始化中 )
      { S7_Templates := "SrcType := Int" } EQ_Contact(in1 := "初始化数据".初始化步骤, in2 := 30)
      Contact( "运动控制数据块".轴初始化错误 )
      Move(in := 90, out1 => "初始化数据".初始化步骤)
   END_RUNG
   // the same network as SCL:
   IF "初始化数据".初始化中 AND ("初始化数据".初始化步骤 = 30) THEN "运动控制数据块".轴初始化按钮 := TRUE; END_IF;
   IF "初始化数据".初始化中 AND ("初始化数据".初始化步骤 = 30) AND "运动控制数据块".轴初始化完成 THEN "初始化数据".初始化步骤 := 40; END_IF;
   IF "初始化数据".初始化中 AND ("初始化数据".初始化步骤 = 30) AND "运动控制数据块".轴初始化错误 THEN "初始化数据".初始化步骤 := 90; END_IF;
END_REGION

REGION Network 8
   RUNG wire#powerrail
      Contact( "初始化数据".初始化中 )
      { S7_Templates := "SrcType := Int" } EQ_Contact(in1 := "初始化数据".初始化步骤, in2 := 40)
      wire#w1
      S_Coil( "初始化数据".初始化完成 )
   END_RUNG
   RUNG wire#w1
      R_Coil( "初始化数据".初始化故障 )
   END_RUNG
   RUNG wire#w1
      R_Coil( "初始化数据".初始化中 )
   END_RUNG
   RUNG wire#w1
      Move(in := 0, out1 => "初始化数据".初始化步骤)
   END_RUNG
   RUNG wire#powerrail
      Contact( "初始化数据".初始化中 )
      { S7_Templates := "SrcType := Int" } EQ_Contact(in1 := "初始化数据".初始化步骤, in2 := 90)
      wire#w2
      S_Coil( "初始化数据".初始化故障 )
   END_RUNG
   RUNG wire#w2
      R_Coil( "初始化数据".初始化中 )
   END_RUNG
   RUNG wire#w2
      Move(in := 0, out1 => "初始化数据".初始化步骤)
   END_RUNG
   // the same network as SCL:
   IF "初始化数据".初始化中 AND ("初始化数据".初始化步骤 = 40) THEN
       "初始化数据".初始化完成 := TRUE;
       "初始化数据".初始化故障 := FALSE;
   END_IF;
   #_w1 := "初始化数据".初始化中 AND ("初始化数据".初始化步骤 = 40);
   IF #_w1 THEN
       "初始化数据".初始化中 := FALSE;
       "初始化数据".初始化步骤 := 0;
   END_IF;
   IF "初始化数据".初始化中 AND ("初始化数据".初始化步骤 = 90) THEN "初始化数据".初始化故障 := TRUE; END_IF;
   #_w2 := "初始化数据".初始化中 AND ("初始化数据".初始化步骤 = 90);
   IF #_w2 THEN
       "初始化数据".初始化中 := FALSE;
       "初始化数据".初始化步骤 := 0;
   END_IF;
END_REGION

REGION Network 9
   RUNG wire#powerrail
      Contact( "状态控制数据".故障状态 )
      R_Coil( "初始化数据".初始化完成 )
   END_RUNG
   // the same network as SCL:
   IF "状态控制数据".故障状态 THEN "初始化数据".初始化完成 := FALSE; END_IF;
END_REGION
END_FUNCTION

FUNCTION "2.状态控制" : Void   // FC22, LAD
{ S7_Optimized_Access := 'TRUE' }
VERSION : 0.1
BEGIN

REGION Network 1: 一站状态判断
   // 故障可加光栅
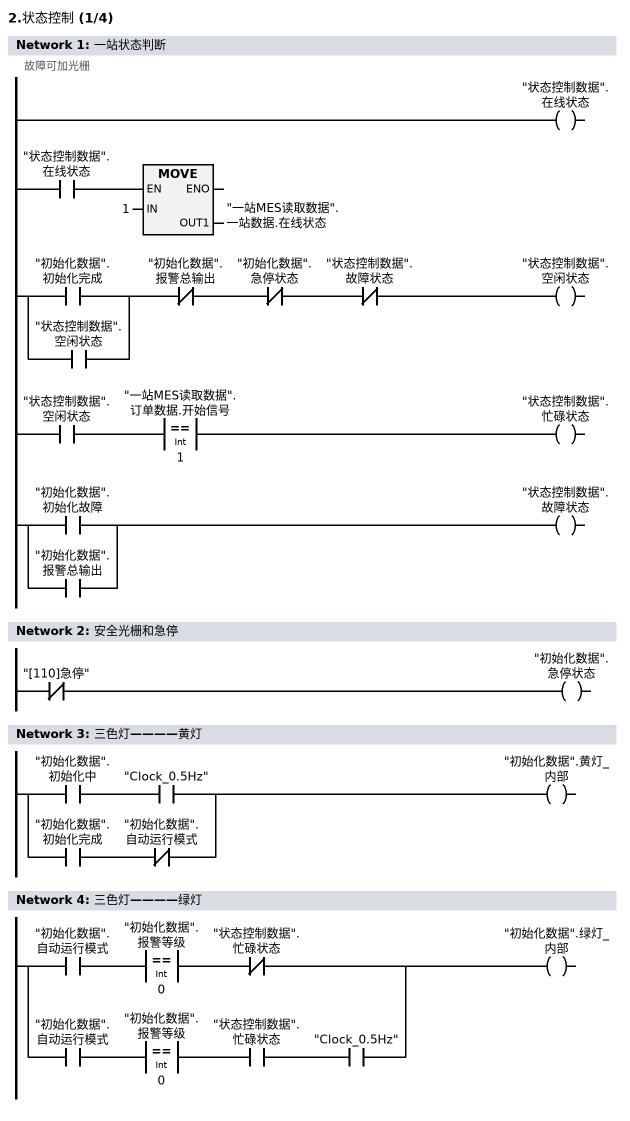
   RUNG wire#powerrail
      Coil( "状态控制数据".在线状态 )
   END_RUNG
   RUNG wire#powerrail
      Contact( "状态控制数据".在线状态 )
      Move(in := 1, out1 => "一站MES读取数据".一站数据.在线状态)
   END_RUNG
   RUNG wire#powerrail
      Contact( "初始化数据".初始化完成 )
      wire#w1
      I_Contact( "初始化数据".报警总输出 )
      I_Contact( "初始化数据".急停状态 )
      I_Contact( "状态控制数据".故障状态 )
      Coil( "状态控制数据".空闲状态 )
   END_RUNG
   RUNG wire#powerrail
      Contact( "状态控制数据".空闲状态 )
   END_RUNG wire#w1
   RUNG wire#powerrail
      Contact( "状态控制数据".空闲状态 )
      { S7_Templates := "SrcType := Int" } EQ_Contact(in1 := "一站MES读取数据".订单数据.开始信号, in2 := 1)
      Coil( "状态控制数据".忙碌状态 )
   END_RUNG
   RUNG wire#powerrail
      Contact( "初始化数据".初始化故障 )
      wire#w2
      Coil( "状态控制数据".故障状态 )
   END_RUNG
   RUNG wire#powerrail
      Contact( "初始化数据".报警总输出 )
   END_RUNG wire#w2
   // the same network as SCL:
   "状态控制数据".在线状态 := TRUE;
   IF "状态控制数据".在线状态 THEN "一站MES读取数据".一站数据.在线状态 := 1; END_IF;
   "状态控制数据".空闲状态 := ("初始化数据".初始化完成 OR "状态控制数据".空闲状态) AND NOT "初始化数据".报警总输出 AND NOT "初始化数据".急停状态 AND NOT "状态控制数据".故障状态;
   "状态控制数据".忙碌状态 := "状态控制数据".空闲状态 AND ("一站MES读取数据".订单数据.开始信号 = 1);
   "状态控制数据".故障状态 := "初始化数据".初始化故障 OR "初始化数据".报警总输出;
END_REGION

REGION Network 2: 安全光栅和急停
   RUNG wire#powerrail
      I_Contact( "[110]急停" )
      Coil( "初始化数据".急停状态 )
   END_RUNG
   // the same network as SCL:
   "初始化数据".急停状态 := NOT "[110]急停";
END_REGION

REGION Network 3: 三色灯————黄灯
   RUNG wire#powerrail
      Contact( "初始化数据".初始化中 )
      Contact( "Clock_0.5Hz" )
      wire#w1
      Coil( "初始化数据".黄灯_内部 )
   END_RUNG
   RUNG wire#powerrail
      Contact( "初始化数据".初始化完成 )
      I_Contact( "初始化数据".自动运行模式 )
   END_RUNG wire#w1
   // the same network as SCL:
   "初始化数据".黄灯_内部 := ("初始化数据".初始化中 AND "Clock_0.5Hz") OR ("初始化数据".初始化完成 AND NOT "初始化数据".自动运行模式);
END_REGION

REGION Network 4: 三色灯————绿灯
   RUNG wire#powerrail
      Contact( "初始化数据".自动运行模式 )
      { S7_Templates := "SrcType := Int" } EQ_Contact(in1 := "初始化数据".报警等级, in2 := 0)
      I_Contact( "状态控制数据".忙碌状态 )
      wire#w1
      Coil( "初始化数据".绿灯_内部 )
   END_RUNG
   RUNG wire#powerrail
      Contact( "初始化数据".自动运行模式 )
      { S7_Templates := "SrcType := Int" } EQ_Contact(in1 := "初始化数据".报警等级, in2 := 0)
      Contact( "状态控制数据".忙碌状态 )
      Contact( "Clock_0.5Hz" )
   END_RUNG wire#w1
   // the same network as SCL:
   "初始化数据".绿灯_内部 := ("初始化数据".自动运行模式 AND ("初始化数据".报警等级 = 0) AND NOT "状态控制数据".忙碌状态) OR ("初始化数据".自动运行模式 AND ("初始化数据".报警等级 = 0) AND "状态控制数据".忙碌状态 AND "Clock_0.5Hz");
END_REGION

REGION Network 5: 三色灯————红灯
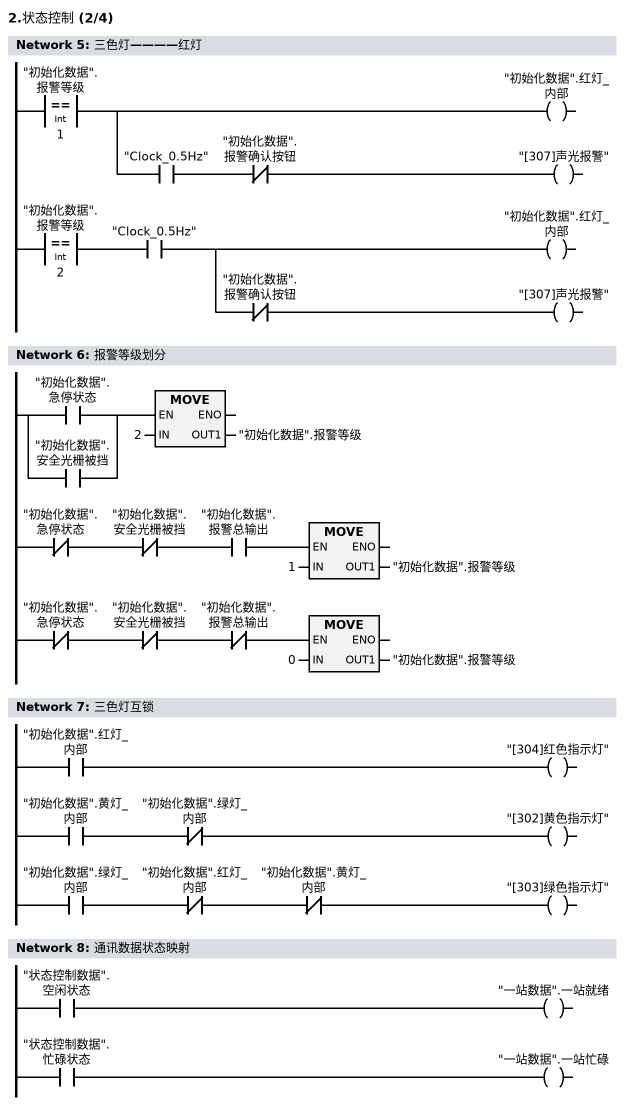
   RUNG wire#powerrail
      { S7_Templates := "SrcType := Int" } EQ_Contact(in1 := "初始化数据".报警等级, in2 := 1)
      wire#w1
      Coil( "初始化数据".红灯_内部 )
   END_RUNG
   RUNG wire#w1
      Contact( "Clock_0.5Hz" )
      I_Contact( "初始化数据".报警确认按钮 )
      Coil( "[307]声光报警" )
   END_RUNG
   RUNG wire#powerrail
      { S7_Templates := "SrcType := Int" } EQ_Contact(in1 := "初始化数据".报警等级, in2 := 2)
      Contact( "Clock_0.5Hz" )
      wire#w2
      Coil( "初始化数据".红灯_内部 )
   END_RUNG
   RUNG wire#w2
      I_Contact( "初始化数据".报警确认按钮 )
      Coil( "[307]声光报警" )
   END_RUNG
   // the same network as SCL:
   "初始化数据".红灯_内部 := "初始化数据".报警等级 = 1;
   "[307]声光报警" := "初始化数据".红灯_内部 AND "Clock_0.5Hz" AND NOT "初始化数据".报警确认按钮;
   "初始化数据".红灯_内部 := ("初始化数据".报警等级 = 2) AND "Clock_0.5Hz";
   "[307]声光报警" := "初始化数据".红灯_内部 AND NOT "初始化数据".报警确认按钮;
END_REGION

REGION Network 6: 报警等级划分
   RUNG wire#powerrail
      Contact( "初始化数据".急停状态 )
      wire#w1
      Move(in := 2, out1 => "初始化数据".报警等级)
   END_RUNG
   RUNG wire#powerrail
      Contact( "初始化数据".安全光栅被挡 )
   END_RUNG wire#w1
   RUNG wire#powerrail
      I_Contact( "初始化数据".急停状态 )
      I_Contact( "初始化数据".安全光栅被挡 )
      Contact( "初始化数据".报警总输出 )
      Move(in := 1, out1 => "初始化数据".报警等级)
   END_RUNG
   RUNG wire#powerrail
      I_Contact( "初始化数据".急停状态 )
      I_Contact( "初始化数据".安全光栅被挡 )
      I_Contact( "初始化数据".报警总输出 )
      Move(in := 0, out1 => "初始化数据".报警等级)
   END_RUNG
   // the same network as SCL:
   IF "初始化数据".急停状态 OR "初始化数据".安全光栅被挡 THEN "初始化数据".报警等级 := 2; END_IF;
   IF NOT "初始化数据".急停状态 AND NOT "初始化数据".安全光栅被挡 AND "初始化数据".报警总输出 THEN "初始化数据".报警等级 := 1; END_IF;
   IF NOT "初始化数据".急停状态 AND NOT "初始化数据".安全光栅被挡 AND NOT "初始化数据".报警总输出 THEN "初始化数据".报警等级 := 0; END_IF;
END_REGION

REGION Network 7: 三色灯互锁
   RUNG wire#powerrail
      Contact( "初始化数据".红灯_内部 )
      Coil( "[304]红色指示灯" )
   END_RUNG
   RUNG wire#powerrail
      Contact( "初始化数据".黄灯_内部 )
      I_Contact( "初始化数据".绿灯_内部 )
      Coil( "[302]黄色指示灯" )
   END_RUNG
   RUNG wire#powerrail
      Contact( "初始化数据".绿灯_内部 )
      I_Contact( "初始化数据".红灯_内部 )
      I_Contact( "初始化数据".黄灯_内部 )
      Coil( "[303]绿色指示灯" )
   END_RUNG
   // the same network as SCL:
   "[304]红色指示灯" := "初始化数据".红灯_内部;
   "[302]黄色指示灯" := "初始化数据".黄灯_内部 AND NOT "初始化数据".绿灯_内部;
   "[303]绿色指示灯" := "初始化数据".绿灯_内部 AND NOT "初始化数据".红灯_内部 AND NOT "初始化数据".黄灯_内部;
END_REGION

REGION Network 8: 通讯数据状态映射
   RUNG wire#powerrail
      Contact( "状态控制数据".空闲状态 )
      Coil( "一站数据".一站就绪 )
   END_RUNG
   RUNG wire#powerrail
      Contact( "状态控制数据".忙碌状态 )
      Coil( "一站数据".一站忙碌 )
   END_RUNG
   // the same network as SCL:
   "一站数据".一站就绪 := "状态控制数据".空闲状态;
   "一站数据".一站忙碌 := "状态控制数据".忙碌状态;
END_REGION

REGION Network 9: MES数据映射
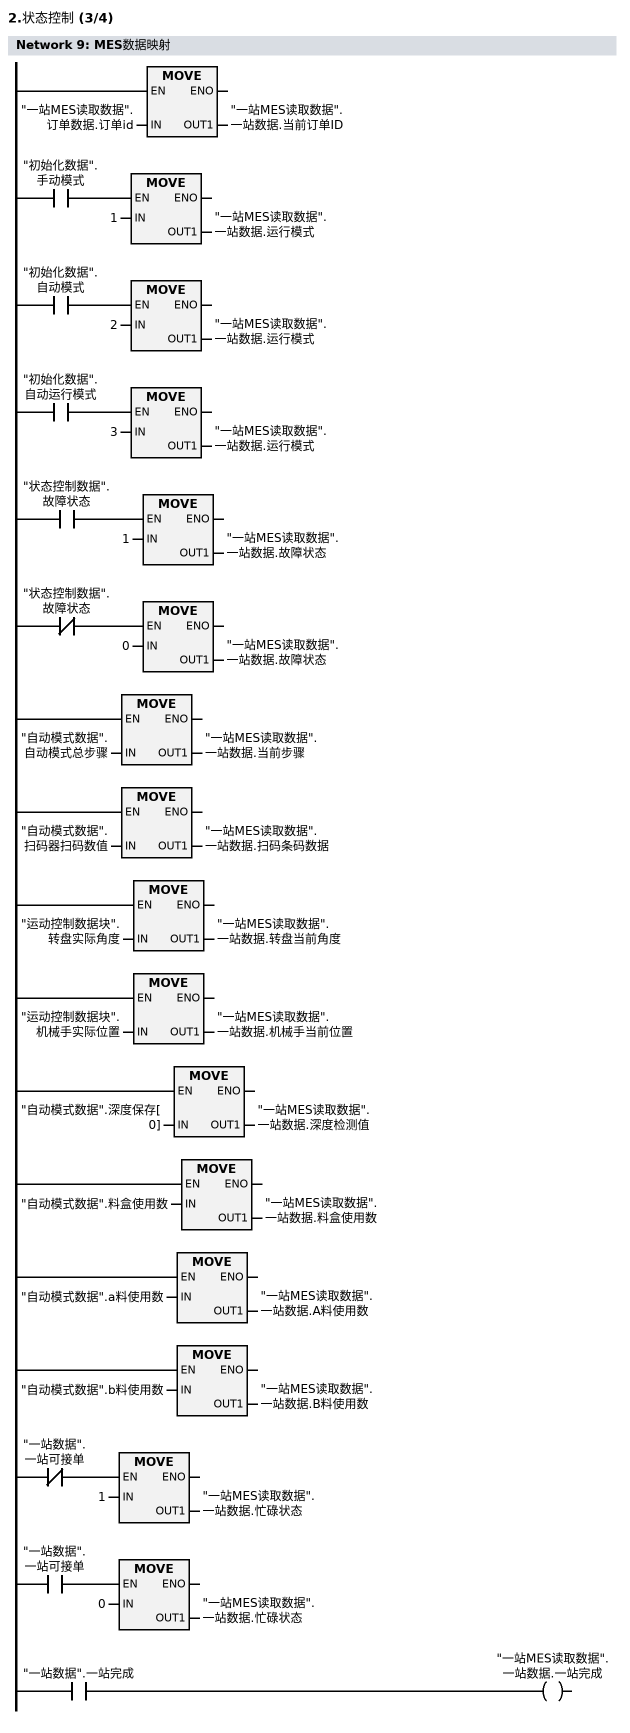
   RUNG wire#powerrail
      Move(in := "一站MES读取数据".订单数据.订单id, out1 => "一站MES读取数据".一站数据.当前订单ID)
   END_RUNG
   RUNG wire#powerrail
      Contact( "初始化数据".手动模式 )
      Move(in := 1, out1 => "一站MES读取数据".一站数据.运行模式)
   END_RUNG
   RUNG wire#powerrail
      Contact( "初始化数据".自动模式 )
      Move(in := 2, out1 => "一站MES读取数据".一站数据.运行模式)
   END_RUNG
   RUNG wire#powerrail
      Contact( "初始化数据".自动运行模式 )
      Move(in := 3, out1 => "一站MES读取数据".一站数据.运行模式)
   END_RUNG
   RUNG wire#powerrail
      Contact( "状态控制数据".故障状态 )
      Move(in := 1, out1 => "一站MES读取数据".一站数据.故障状态)
   END_RUNG
   RUNG wire#powerrail
      I_Contact( "状态控制数据".故障状态 )
      Move(in := 0, out1 => "一站MES读取数据".一站数据.故障状态)
   END_RUNG
   RUNG wire#powerrail
      Move(in := "自动模式数据".自动模式总步骤, out1 => "一站MES读取数据".一站数据.当前步骤)
   END_RUNG
   RUNG wire#powerrail
      Move(in := "自动模式数据".扫码器扫码数值, out1 => "一站MES读取数据".一站数据.扫码条码数据)
   END_RUNG
   RUNG wire#powerrail
      Move(in := "运动控制数据块".转盘实际角度, out1 => "一站MES读取数据".一站数据.转盘当前角度)
   END_RUNG
   RUNG wire#powerrail
      Move(in := "运动控制数据块".机械手实际位置, out1 => "一站MES读取数据".一站数据.机械手当前位置)
   END_RUNG
   RUNG wire#powerrail
      Move(in := "自动模式数据".深度保存[0], out1 => "一站MES读取数据".一站数据.深度检测值)
   END_RUNG
   RUNG wire#powerrail
      Move(in := "自动模式数据".料盒使用数, out1 => "一站MES读取数据".一站数据.料盒使用数)
   END_RUNG
   RUNG wire#powerrail
      Move(in := "自动模式数据".a料使用数, out1 => "一站MES读取数据".一站数据.A料使用数)
   END_RUNG
   RUNG wire#powerrail
      Move(in := "自动模式数据".b料使用数, out1 => "一站MES读取数据".一站数据.B料使用数)
   END_RUNG
   RUNG wire#powerrail
      I_Contact( "一站数据".一站可接单 )
      Move(in := 1, out1 => "一站MES读取数据".一站数据.忙碌状态)
   END_RUNG
   RUNG wire#powerrail
      Contact( "一站数据".一站可接单 )
      Move(in := 0, out1 => "一站MES读取数据".一站数据.忙碌状态)
   END_RUNG
   RUNG wire#powerrail
      Contact( "一站数据".一站完成 )
      Coil( "一站MES读取数据".一站数据.一站完成 )
   END_RUNG
   // the same network as SCL:
   "一站MES读取数据".一站数据.当前订单ID := "一站MES读取数据".订单数据.订单id;
   IF "初始化数据".手动模式 THEN "一站MES读取数据".一站数据.运行模式 := 1; END_IF;
   IF "初始化数据".自动模式 THEN "一站MES读取数据".一站数据.运行模式 := 2; END_IF;
   IF "初始化数据".自动运行模式 THEN "一站MES读取数据".一站数据.运行模式 := 3; END_IF;
   IF "状态控制数据".故障状态 THEN "一站MES读取数据".一站数据.故障状态 := 1; END_IF;
   IF NOT "状态控制数据".故障状态 THEN "一站MES读取数据".一站数据.故障状态 := 0; END_IF;
   "一站MES读取数据".一站数据.当前步骤 := "自动模式数据".自动模式总步骤;
   "一站MES读取数据".一站数据.扫码条码数据 := "自动模式数据".扫码器扫码数值;
   "一站MES读取数据".一站数据.转盘当前角度 := "运动控制数据块".转盘实际角度;
   "一站MES读取数据".一站数据.机械手当前位置 := "运动控制数据块".机械手实际位置;
   "一站MES读取数据".一站数据.深度检测值 := "自动模式数据".深度保存[0];
   "一站MES读取数据".一站数据.料盒使用数 := "自动模式数据".料盒使用数;
   "一站MES读取数据".一站数据.A料使用数 := "自动模式数据".a料使用数;
   "一站MES读取数据".一站数据.B料使用数 := "自动模式数据".b料使用数;
   IF NOT "一站数据".一站可接单 THEN "一站MES读取数据".一站数据.忙碌状态 := 1; END_IF;
   IF "一站数据".一站可接单 THEN "一站MES读取数据".一站数据.忙碌状态 := 0; END_IF;
   "一站MES读取数据".一站数据.一站完成 := "一站数据".一站完成;
END_REGION

REGION Network 10
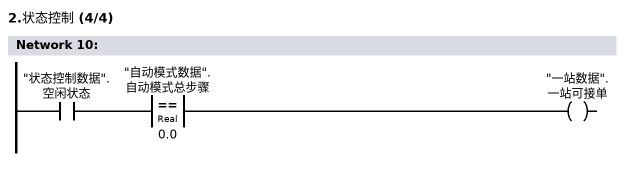
   RUNG wire#powerrail
      Contact( "状态控制数据".空闲状态 )
      { S7_Templates := "SrcType := Real" } EQ_Contact(in1 := "自动模式数据".自动模式总步骤, in2 := 0.0)
      Coil( "一站数据".一站可接单 )
   END_RUNG
   // the same network as SCL:
   "一站数据".一站可接单 := "状态控制数据".空闲状态 AND ("自动模式数据".自动模式总步骤 = 0.0);
END_REGION
END_FUNCTION

ORGANIZATION_BLOCK "Main"   // OB1, LAD, ProgramCycle
TITLE = "Main Program Sweep (Cycle)"
{ S7_Optimized_Access := 'TRUE' }
VERSION : 0.1
// 做MES，MES做完修产线的小问题，还有HMI
   VAR_INPUT
      Initial_Call : Bool;   // Initial call of this OB
      Remanence : Bool;   // =True, if remanent data are available
   END_VAR
   VAR_TEMP   // added for the SCL form of the ladder/FBD networks
      _w1 : Bool;
      _w2 : Bool;
      _w3 : Bool;
      _w4 : Bool;
   END_VAR
BEGIN

REGION Network 1: 自动模式
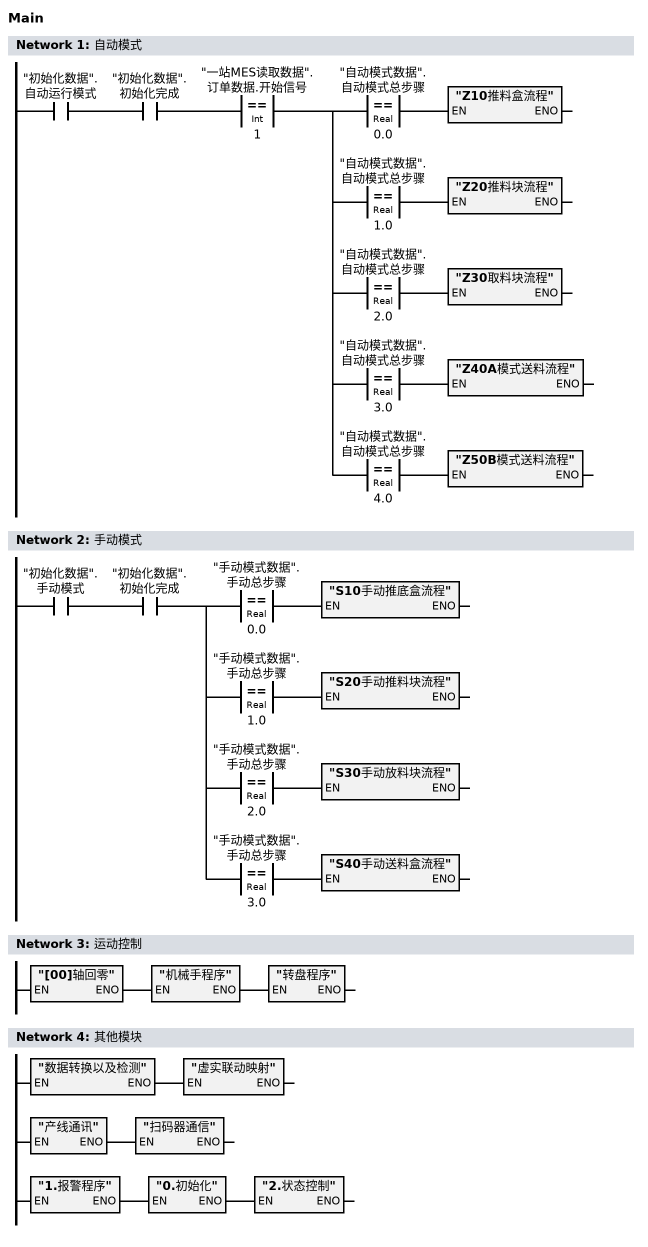
   RUNG wire#powerrail
      Contact( "初始化数据".自动运行模式 )
      Contact( "初始化数据".初始化完成 )
      { S7_Templates := "SrcType := Int" } EQ_Contact(in1 := "一站MES读取数据".订单数据.开始信号, in2 := 1)
      wire#w1
      { S7_Templates := "SrcType := Real" } EQ_Contact(in1 := "自动模式数据".自动模式总步骤, in2 := 0.0)
      "Z10推料盒流程"()
   END_RUNG
   RUNG wire#w1
      { S7_Templates := "SrcType := Real" } EQ_Contact(in1 := "自动模式数据".自动模式总步骤, in2 := 1.0)
      "Z20推料块流程"()
   END_RUNG
   RUNG wire#w1
      { S7_Templates := "SrcType := Real" } EQ_Contact(in1 := "自动模式数据".自动模式总步骤, in2 := 2.0)
      "Z30取料块流程"()
   END_RUNG
   RUNG wire#w1
      { S7_Templates := "SrcType := Real" } EQ_Contact(in1 := "自动模式数据".自动模式总步骤, in2 := 3.0)
      "Z40A模式送料流程"()
   END_RUNG
   RUNG wire#w1
      { S7_Templates := "SrcType := Real" } EQ_Contact(in1 := "自动模式数据".自动模式总步骤, in2 := 4.0)
      "Z50B模式送料流程"()
   END_RUNG
   // the same network as SCL:
   #_w1 := "初始化数据".自动运行模式 AND "初始化数据".初始化完成 AND ("一站MES读取数据".订单数据.开始信号 = 1);
   IF #_w1 AND ("自动模式数据".自动模式总步骤 = 0.0) THEN "Z10推料盒流程"(); END_IF;
   IF #_w1 AND ("自动模式数据".自动模式总步骤 = 1.0) THEN "Z20推料块流程"(); END_IF;
   IF #_w1 AND ("自动模式数据".自动模式总步骤 = 2.0) THEN "Z30取料块流程"(); END_IF;
   IF #_w1 AND ("自动模式数据".自动模式总步骤 = 3.0) THEN "Z40A模式送料流程"(); END_IF;
   IF #_w1 AND ("自动模式数据".自动模式总步骤 = 4.0) THEN "Z50B模式送料流程"(); END_IF;
END_REGION

REGION Network 2: 手动模式
   RUNG wire#powerrail
      Contact( "初始化数据".手动模式 )
      Contact( "初始化数据".初始化完成 )
      wire#w1
      { S7_Templates := "SrcType := Real" } EQ_Contact(in1 := "手动模式数据".手动总步骤, in2 := 0.0)
      "S10手动推底盒流程"()
   END_RUNG
   RUNG wire#w1
      { S7_Templates := "SrcType := Real" } EQ_Contact(in1 := "手动模式数据".手动总步骤, in2 := 1.0)
      "S20手动推料块流程"()
   END_RUNG
   RUNG wire#w1
      { S7_Templates := "SrcType := Real" } EQ_Contact(in1 := "手动模式数据".手动总步骤, in2 := 2.0)
      "S30手动放料块流程"()
   END_RUNG
   RUNG wire#w1
      { S7_Templates := "SrcType := Real" } EQ_Contact(in1 := "手动模式数据".手动总步骤, in2 := 3.0)
      "S40手动送料盒流程"()
   END_RUNG
   // the same network as SCL:
   #_w1 := "初始化数据".手动模式 AND "初始化数据".初始化完成;
   IF #_w1 AND ("手动模式数据".手动总步骤 = 0.0) THEN "S10手动推底盒流程"(); END_IF;
   IF #_w1 AND ("手动模式数据".手动总步骤 = 1.0) THEN "S20手动推料块流程"(); END_IF;
   IF #_w1 AND ("手动模式数据".手动总步骤 = 2.0) THEN "S30手动放料块流程"(); END_IF;
   IF #_w1 AND ("手动模式数据".手动总步骤 = 3.0) THEN "S40手动送料盒流程"(); END_IF;
END_REGION

REGION Network 3: 运动控制
   RUNG wire#powerrail
      "[00]轴回零"()
      "机械手程序"()
      "转盘程序"()
   END_RUNG
   // the same network as SCL:
   "[00]轴回零"(ENO => #_w1);
   "机械手程序"(EN := #_w1, ENO => #_w2);
   IF #_w2 THEN "转盘程序"(); END_IF;
END_REGION

REGION Network 4: 其他模块
   RUNG wire#powerrail
      "数据转换以及检测"()
      "虚实联动映射"()
   END_RUNG
   RUNG wire#powerrail
      "产线通讯"()
      "扫码器通信"()
   END_RUNG
   RUNG wire#powerrail
      "1.报警程序"()
      "0.初始化"()
      "2.状态控制"()
   END_RUNG
   // the same network as SCL:
   "数据转换以及检测"(ENO => #_w1);
   IF #_w1 THEN "虚实联动映射"(); END_IF;
   "产线通讯"(ENO => #_w2);
   IF #_w2 THEN "扫码器通信"(); END_IF;
   "1.报警程序"(ENO => #_w3);
   "0.初始化"(EN := #_w3, ENO => #_w4);
   IF #_w4 THEN "2.状态控制"(); END_IF;
END_REGION
END_ORGANIZATION_BLOCK

// folder: 手动模式

FUNCTION "S10手动推底盒流程" : Void   // FC2, LAD
TITLE = 该流程将底盒推出到转盘
{ S7_Optimized_Access := 'TRUE' }
VERSION : 0.1
   VAR_TEMP   // added for the SCL form of the ladder/FBD networks
      _w1 : Bool;
      _w2 : Bool;
   END_VAR
BEGIN

REGION Network 1: 气缸推出
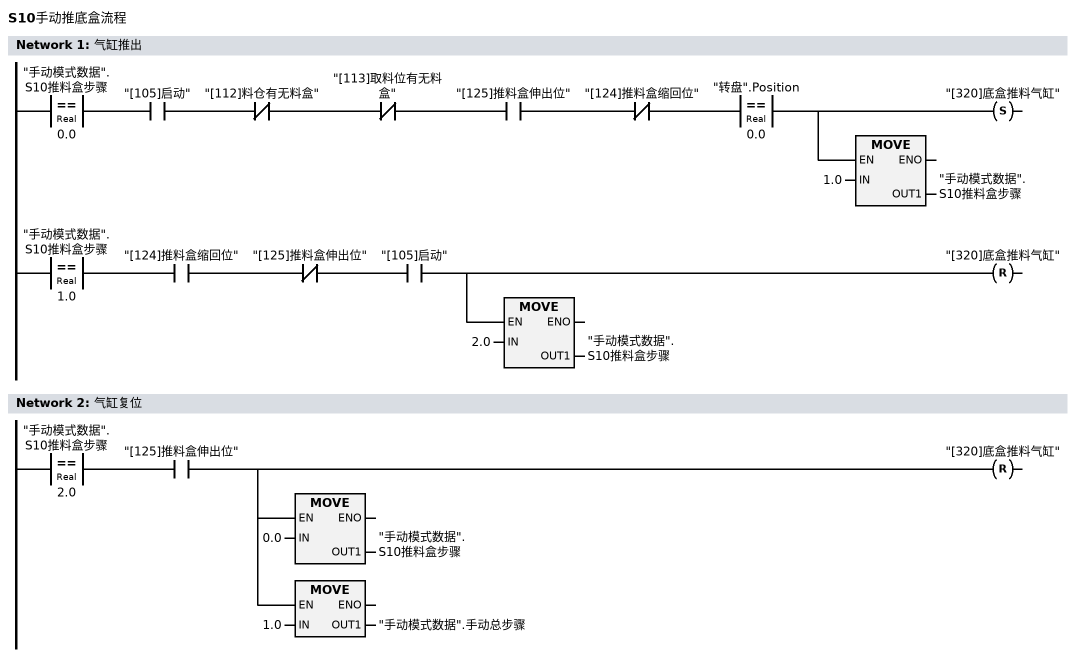
   RUNG wire#powerrail
      { S7_Templates := "SrcType := Real" } EQ_Contact(in1 := "手动模式数据".S10推料盒步骤, in2 := 0.0)
      Contact( "[105]启动" )
      I_Contact( "[112]料仓有无料盒" )
      I_Contact( "[113]取料位有无料盒" )
      Contact( "[125]推料盒伸出位" )
      I_Contact( "[124]推料盒缩回位" )
      { S7_Templates := "SrcType := Real" } EQ_Contact(in1 := "转盘".Position, in2 := 0.0)
      wire#w1
      S_Coil( "[320]底盒推料气缸" )
   END_RUNG
   RUNG wire#w1
      Move(in := 1.0, out1 => "手动模式数据".S10推料盒步骤)
   END_RUNG
   RUNG wire#powerrail
      { S7_Templates := "SrcType := Real" } EQ_Contact(in1 := "手动模式数据".S10推料盒步骤, in2 := 1.0)
      Contact( "[124]推料盒缩回位" )
      I_Contact( "[125]推料盒伸出位" )
      Contact( "[105]启动" )
      wire#w2
      R_Coil( "[320]底盒推料气缸" )
   END_RUNG
   RUNG wire#w2
      Move(in := 2.0, out1 => "手动模式数据".S10推料盒步骤)
   END_RUNG
   // the same network as SCL:
   #_w1 := ("手动模式数据".S10推料盒步骤 = 0.0) AND "[105]启动" AND NOT "[112]料仓有无料盒" AND NOT "[113]取料位有无料盒" AND "[125]推料盒伸出位" AND NOT "[124]推料盒缩回位" AND ("转盘".Position = 0.0);
   IF #_w1 THEN
       "[320]底盒推料气缸" := TRUE;
       "手动模式数据".S10推料盒步骤 := 1.0;
   END_IF;
   #_w2 := ("手动模式数据".S10推料盒步骤 = 1.0) AND "[124]推料盒缩回位" AND NOT "[125]推料盒伸出位" AND "[105]启动";
   IF #_w2 THEN
       "[320]底盒推料气缸" := FALSE;
       "手动模式数据".S10推料盒步骤 := 2.0;
   END_IF;
END_REGION

REGION Network 2: 气缸复位
   RUNG wire#powerrail
      { S7_Templates := "SrcType := Real" } EQ_Contact(in1 := "手动模式数据".S10推料盒步骤, in2 := 2.0)
      Contact( "[125]推料盒伸出位" )
      wire#w1
      R_Coil( "[320]底盒推料气缸" )
   END_RUNG
   RUNG wire#w1
      Move(in := 0.0, out1 => "手动模式数据".S10推料盒步骤)
   END_RUNG
   RUNG wire#w1
      Move(in := 1.0, out1 => "手动模式数据".手动总步骤)
   END_RUNG
   // the same network as SCL:
   #_w1 := ("手动模式数据".S10推料盒步骤 = 2.0) AND "[125]推料盒伸出位";
   IF #_w1 THEN
       "[320]底盒推料气缸" := FALSE;
       "手动模式数据".S10推料盒步骤 := 0.0;
       "手动模式数据".手动总步骤 := 1.0;
   END_IF;
END_REGION
END_FUNCTION

FUNCTION "S20手动推料块流程" : Void   // FC3, LAD
TITLE = 该流程从AB库推出料块
{ S7_Optimized_Access := 'TRUE' }
VERSION : 0.1
   VAR_TEMP   // added for the SCL form of the ladder/FBD networks
      _w1 : Bool;
      _w2 : Bool;
      _w3 : Bool;
   END_VAR
BEGIN

REGION Network 1
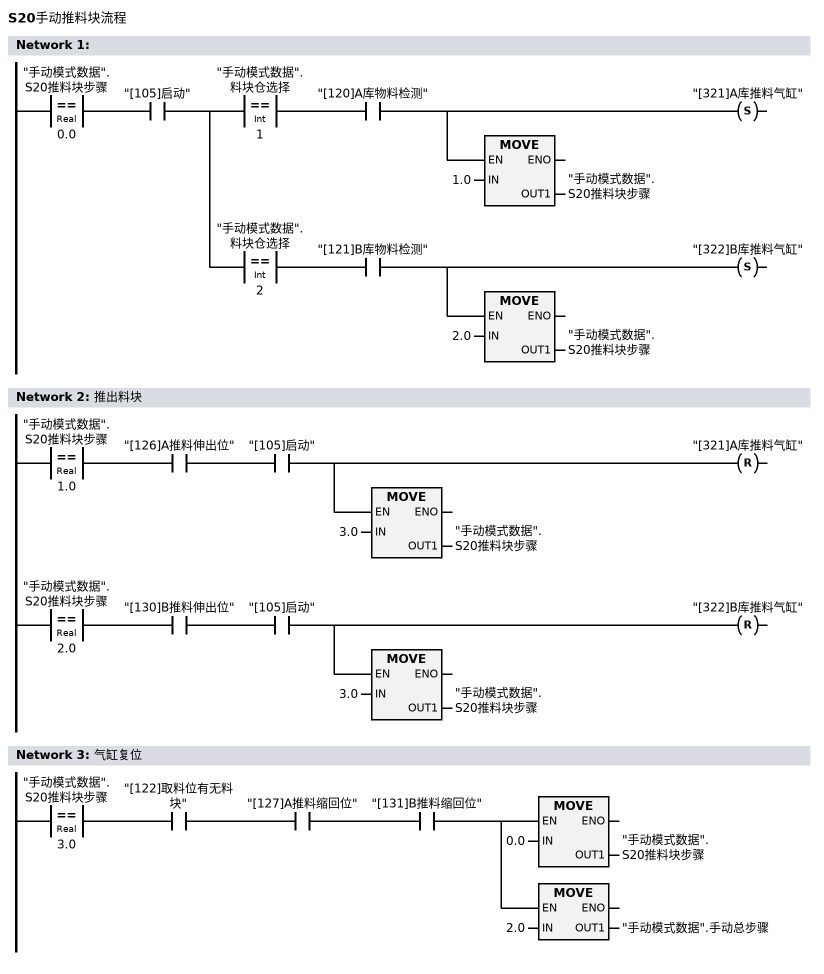
   RUNG wire#powerrail
      { S7_Templates := "SrcType := Real" } EQ_Contact(in1 := "手动模式数据".S20推料块步骤, in2 := 0.0)
      Contact( "[105]启动" )
      wire#w1
      { S7_Templates := "SrcType := Int" } EQ_Contact(in1 := "手动模式数据".料块仓选择, in2 := 1)
      Contact( "[120]A库物料检测" )
      wire#w2
      S_Coil( "[321]A库推料气缸" )
   END_RUNG
   RUNG wire#w2
      Move(in := 1.0, out1 => "手动模式数据".S20推料块步骤)
   END_RUNG
   RUNG wire#w1
      { S7_Templates := "SrcType := Int" } EQ_Contact(in1 := "手动模式数据".料块仓选择, in2 := 2)
      Contact( "[121]B库物料检测" )
      wire#w3
      S_Coil( "[322]B库推料气缸" )
   END_RUNG
   RUNG wire#w3
      Move(in := 2.0, out1 => "手动模式数据".S20推料块步骤)
   END_RUNG
   // the same network as SCL:
   #_w1 := ("手动模式数据".S20推料块步骤 = 0.0) AND "[105]启动";
   #_w2 := #_w1 AND ("手动模式数据".料块仓选择 = 1) AND "[120]A库物料检测";
   IF #_w2 THEN
       "[321]A库推料气缸" := TRUE;
       "手动模式数据".S20推料块步骤 := 1.0;
   END_IF;
   #_w3 := #_w1 AND ("手动模式数据".料块仓选择 = 2) AND "[121]B库物料检测";
   IF #_w3 THEN
       "[322]B库推料气缸" := TRUE;
       "手动模式数据".S20推料块步骤 := 2.0;
   END_IF;
END_REGION

REGION Network 2: 推出料块
   RUNG wire#powerrail
      { S7_Templates := "SrcType := Real" } EQ_Contact(in1 := "手动模式数据".S20推料块步骤, in2 := 1.0)
      Contact( "[126]A推料伸出位" )
      Contact( "[105]启动" )
      wire#w1
      R_Coil( "[321]A库推料气缸" )
   END_RUNG
   RUNG wire#w1
      Move(in := 3.0, out1 => "手动模式数据".S20推料块步骤)
   END_RUNG
   RUNG wire#powerrail
      { S7_Templates := "SrcType := Real" } EQ_Contact(in1 := "手动模式数据".S20推料块步骤, in2 := 2.0)
      Contact( "[130]B推料伸出位" )
      Contact( "[105]启动" )
      wire#w2
      R_Coil( "[322]B库推料气缸" )
   END_RUNG
   RUNG wire#w2
      Move(in := 3.0, out1 => "手动模式数据".S20推料块步骤)
   END_RUNG
   // the same network as SCL:
   #_w1 := ("手动模式数据".S20推料块步骤 = 1.0) AND "[126]A推料伸出位" AND "[105]启动";
   IF #_w1 THEN
       "[321]A库推料气缸" := FALSE;
       "手动模式数据".S20推料块步骤 := 3.0;
   END_IF;
   #_w2 := ("手动模式数据".S20推料块步骤 = 2.0) AND "[130]B推料伸出位" AND "[105]启动";
   IF #_w2 THEN
       "[322]B库推料气缸" := FALSE;
       "手动模式数据".S20推料块步骤 := 3.0;
   END_IF;
END_REGION

REGION Network 3: 气缸复位
   RUNG wire#powerrail
      { S7_Templates := "SrcType := Real" } EQ_Contact(in1 := "手动模式数据".S20推料块步骤, in2 := 3.0)
      Contact( "[122]取料位有无料块" )
      Contact( "[127]A推料缩回位" )
      Contact( "[131]B推料缩回位" )
      wire#w1
      Move(in := 0.0, out1 => "手动模式数据".S20推料块步骤)
   END_RUNG
   RUNG wire#w1
      Move(in := 2.0, out1 => "手动模式数据".手动总步骤)
   END_RUNG
   // the same network as SCL:
   #_w1 := ("手动模式数据".S20推料块步骤 = 3.0) AND "[122]取料位有无料块" AND "[127]A推料缩回位" AND "[131]B推料缩回位";
   IF #_w1 THEN
       "手动模式数据".S20推料块步骤 := 0.0;
       "手动模式数据".手动总步骤 := 2.0;
   END_IF;
END_REGION
END_FUNCTION

FUNCTION "S40手动送料盒流程" : Void   // FC6, LAD
{ S7_Optimized_Access := 'TRUE' }
VERSION : 0.1
// 深度检测后夹到第二站
   VAR_TEMP   // added for the SCL form of the ladder/FBD networks
      _w1 : Bool;
      _w2 : Bool;
   END_VAR
BEGIN

REGION Network 1
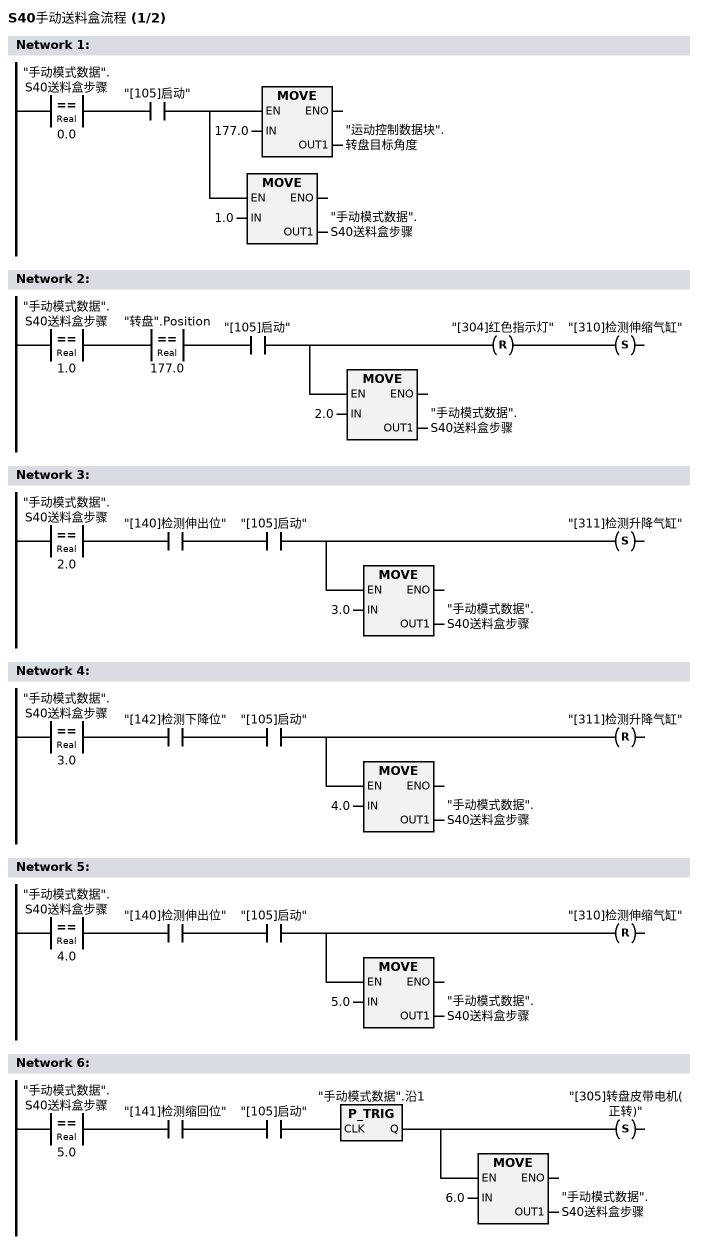
   RUNG wire#powerrail
      { S7_Templates := "SrcType := Real" } EQ_Contact(in1 := "手动模式数据".S40送料盒步骤, in2 := 0.0)
      Contact( "[105]启动" )
      wire#w1
      Move(in := 177.0, out1 => "运动控制数据块".转盘目标角度)
   END_RUNG
   RUNG wire#w1
      Move(in := 1.0, out1 => "手动模式数据".S40送料盒步骤)
   END_RUNG
   // the same network as SCL:
   IF ("手动模式数据".S40送料盒步骤 = 0.0) AND "[105]启动" THEN
       "运动控制数据块".转盘目标角度 := 177.0;
       "手动模式数据".S40送料盒步骤 := 1.0;
   END_IF;
END_REGION

REGION Network 2
   RUNG wire#powerrail
      { S7_Templates := "SrcType := Real" } EQ_Contact(in1 := "手动模式数据".S40送料盒步骤, in2 := 1.0)
      { S7_Templates := "SrcType := Real" } EQ_Contact(in1 := "转盘".Position, in2 := 177.0)
      Contact( "[105]启动" )
      wire#w1
      R_Coil( "[304]红色指示灯" )
      S_Coil( "[310]检测伸缩气缸" )
   END_RUNG
   RUNG wire#w1
      Move(in := 2.0, out1 => "手动模式数据".S40送料盒步骤)
   END_RUNG
   // the same network as SCL:
   #_w1 := ("手动模式数据".S40送料盒步骤 = 1.0) AND ("转盘".Position = 177.0) AND "[105]启动";
   IF #_w1 THEN
       "[304]红色指示灯" := FALSE;
       "[310]检测伸缩气缸" := TRUE;
       "手动模式数据".S40送料盒步骤 := 2.0;
   END_IF;
END_REGION

REGION Network 3
   RUNG wire#powerrail
      { S7_Templates := "SrcType := Real" } EQ_Contact(in1 := "手动模式数据".S40送料盒步骤, in2 := 2.0)
      Contact( "[140]检测伸出位" )
      Contact( "[105]启动" )
      wire#w1
      S_Coil( "[311]检测升降气缸" )
   END_RUNG
   RUNG wire#w1
      Move(in := 3.0, out1 => "手动模式数据".S40送料盒步骤)
   END_RUNG
   // the same network as SCL:
   #_w1 := ("手动模式数据".S40送料盒步骤 = 2.0) AND "[140]检测伸出位" AND "[105]启动";
   IF #_w1 THEN
       "[311]检测升降气缸" := TRUE;
       "手动模式数据".S40送料盒步骤 := 3.0;
   END_IF;
END_REGION

REGION Network 4
   RUNG wire#powerrail
      { S7_Templates := "SrcType := Real" } EQ_Contact(in1 := "手动模式数据".S40送料盒步骤, in2 := 3.0)
      Contact( "[142]检测下降位" )
      Contact( "[105]启动" )
      wire#w1
      R_Coil( "[311]检测升降气缸" )
   END_RUNG
   RUNG wire#w1
      Move(in := 4.0, out1 => "手动模式数据".S40送料盒步骤)
   END_RUNG
   // the same network as SCL:
   #_w1 := ("手动模式数据".S40送料盒步骤 = 3.0) AND "[142]检测下降位" AND "[105]启动";
   IF #_w1 THEN
       "[311]检测升降气缸" := FALSE;
       "手动模式数据".S40送料盒步骤 := 4.0;
   END_IF;
END_REGION

REGION Network 5
   RUNG wire#powerrail
      { S7_Templates := "SrcType := Real" } EQ_Contact(in1 := "手动模式数据".S40送料盒步骤, in2 := 4.0)
      Contact( "[140]检测伸出位" )
      Contact( "[105]启动" )
      wire#w1
      R_Coil( "[310]检测伸缩气缸" )
   END_RUNG
   RUNG wire#w1
      Move(in := 5.0, out1 => "手动模式数据".S40送料盒步骤)
   END_RUNG
   // the same network as SCL:
   #_w1 := ("手动模式数据".S40送料盒步骤 = 4.0) AND "[140]检测伸出位" AND "[105]启动";
   IF #_w1 THEN
       "[310]检测伸缩气缸" := FALSE;
       "手动模式数据".S40送料盒步骤 := 5.0;
   END_IF;
END_REGION

REGION Network 6
   RUNG wire#powerrail
      { S7_Templates := "SrcType := Real" } EQ_Contact(in1 := "手动模式数据".S40送料盒步骤, in2 := 5.0)
      Contact( "[141]检测缩回位" )
      Contact( "[105]启动" )
      P_Trig( "手动模式数据".沿1 )
      wire#w1
      S_Coil( "[305]转盘皮带电机(正转)" )
   END_RUNG
   RUNG wire#w1
      Move(in := 6.0, out1 => "手动模式数据".S40送料盒步骤)
   END_RUNG
   // the same network as SCL:
   #_w1 := ("手动模式数据".S40送料盒步骤 = 5.0) AND "[141]检测缩回位" AND "[105]启动";
   #_w2 := #_w1 AND NOT "手动模式数据".沿1;   // rising edge
   "手动模式数据".沿1 := #_w1;
   IF #_w2 THEN
       "[305]转盘皮带电机(正转)" := TRUE;
       "手动模式数据".S40送料盒步骤 := 6.0;
   END_IF;
END_REGION

REGION Network 7
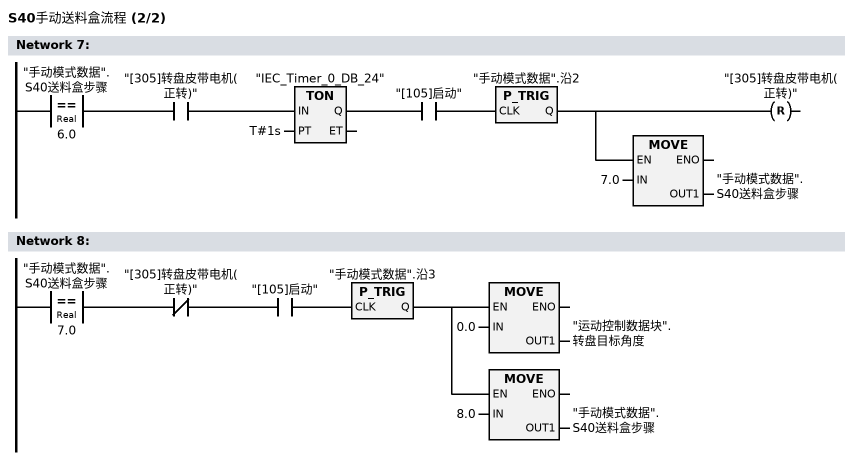
   "IEC_Timer_0_DB_24".TON(IN := ("手动模式数据".S40送料盒步骤 = 6.0) AND "[305]转盘皮带电机(正转)", PT := T#1s);
   #_w1 := "IEC_Timer_0_DB_24".Q AND "[105]启动";
   #_w2 := #_w1 AND NOT "手动模式数据".沿2;   // rising edge
   "手动模式数据".沿2 := #_w1;
   IF #_w2 THEN
       "[305]转盘皮带电机(正转)" := FALSE;
       "手动模式数据".S40送料盒步骤 := 7.0;
   END_IF;
END_REGION

REGION Network 8
   RUNG wire#powerrail
      { S7_Templates := "SrcType := Real" } EQ_Contact(in1 := "手动模式数据".S40送料盒步骤, in2 := 7.0)
      I_Contact( "[305]转盘皮带电机(正转)" )
      Contact( "[105]启动" )
      P_Trig( "手动模式数据".沿3 )
      wire#w1
      Move(in := 0.0, out1 => "运动控制数据块".转盘目标角度)
   END_RUNG
   RUNG wire#w1
      Move(in := 8.0, out1 => "手动模式数据".S40送料盒步骤)
   END_RUNG
   // the same network as SCL:
   #_w1 := ("手动模式数据".S40送料盒步骤 = 7.0) AND NOT "[305]转盘皮带电机(正转)" AND "[105]启动";
   #_w2 := #_w1 AND NOT "手动模式数据".沿3;   // rising edge
   "手动模式数据".沿3 := #_w1;
   IF #_w2 THEN
       "运动控制数据块".转盘目标角度 := 0.0;
       "手动模式数据".S40送料盒步骤 := 8.0;
   END_IF;
END_REGION
END_FUNCTION

FUNCTION "S30手动放料块流程" : Void   // FC7, LAD
TITLE = 该流程将料块放到底盒
{ S7_Optimized_Access := 'TRUE' }
VERSION : 0.1
   VAR_TEMP   // added for the SCL form of the ladder/FBD networks
      _w1 : Bool;
      _w2 : Bool;
      _w3 : Bool;
   END_VAR
BEGIN

REGION Network 1: 吸取料块
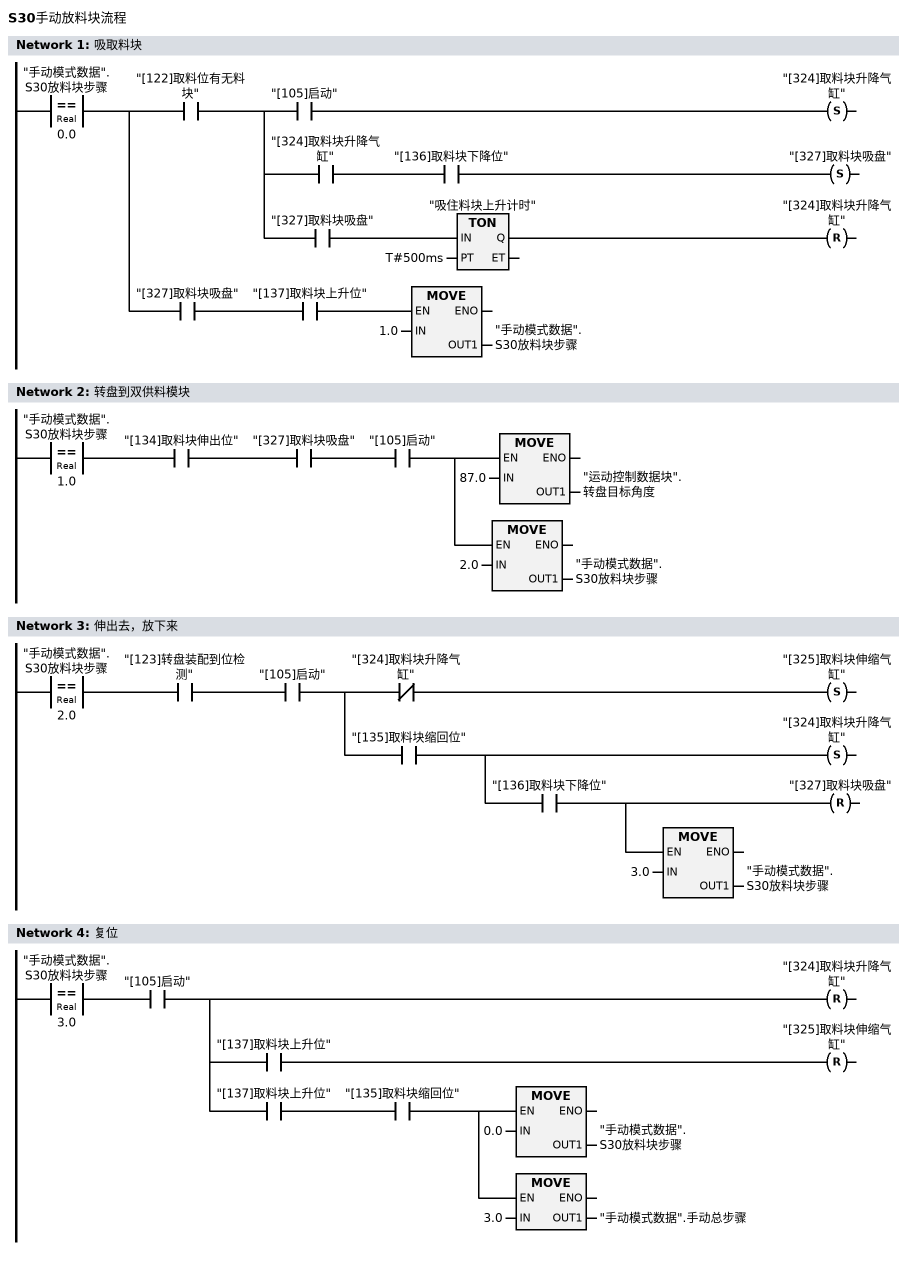
   #_w1 := "手动模式数据".S30放料块步骤 = 0.0;
   #_w2 := #_w1 AND "[122]取料位有无料块";
   IF #_w2 AND "[105]启动" THEN "[324]取料块升降气缸" := TRUE; END_IF;
   IF #_w2 AND "[324]取料块升降气缸" AND "[136]取料块下降位" THEN "[327]取料块吸盘" := TRUE; END_IF;
   "吸住料块上升计时".TON(IN := #_w2 AND "[327]取料块吸盘", PT := T#500ms);
   IF "吸住料块上升计时".Q THEN "[324]取料块升降气缸" := FALSE; END_IF;
   IF #_w1 AND "[327]取料块吸盘" AND "[137]取料块上升位" THEN "手动模式数据".S30放料块步骤 := 1.0; END_IF;
END_REGION

REGION Network 2: 转盘到双供料模块
   RUNG wire#powerrail
      { S7_Templates := "SrcType := Real" } EQ_Contact(in1 := "手动模式数据".S30放料块步骤, in2 := 1.0)
      Contact( "[134]取料块伸出位" )
      Contact( "[327]取料块吸盘" )
      Contact( "[105]启动" )
      wire#w1
      Move(in := 87.0, out1 => "运动控制数据块".转盘目标角度)
   END_RUNG
   RUNG wire#w1
      Move(in := 2.0, out1 => "手动模式数据".S30放料块步骤)
   END_RUNG
   // the same network as SCL:
   IF ("手动模式数据".S30放料块步骤 = 1.0) AND "[134]取料块伸出位" AND "[327]取料块吸盘" AND "[105]启动" THEN
       "运动控制数据块".转盘目标角度 := 87.0;
       "手动模式数据".S30放料块步骤 := 2.0;
   END_IF;
END_REGION

REGION Network 3: 伸出去，放下来
   RUNG wire#powerrail
      { S7_Templates := "SrcType := Real" } EQ_Contact(in1 := "手动模式数据".S30放料块步骤, in2 := 2.0)
      Contact( "[123]转盘装配到位检测" )
      Contact( "[105]启动" )
      wire#w1
      I_Contact( "[324]取料块升降气缸" )
      S_Coil( "[325]取料块伸缩气缸" )
   END_RUNG
   RUNG wire#w1
      Contact( "[135]取料块缩回位" )
      wire#w2
      S_Coil( "[324]取料块升降气缸" )
   END_RUNG
   RUNG wire#w2
      Contact( "[136]取料块下降位" )
      wire#w3
      R_Coil( "[327]取料块吸盘" )
   END_RUNG
   RUNG wire#w3
      Move(in := 3.0, out1 => "手动模式数据".S30放料块步骤)
   END_RUNG
   // the same network as SCL:
   #_w1 := ("手动模式数据".S30放料块步骤 = 2.0) AND "[123]转盘装配到位检测" AND "[105]启动";
   IF #_w1 AND NOT "[324]取料块升降气缸" THEN "[325]取料块伸缩气缸" := TRUE; END_IF;
   #_w2 := #_w1 AND "[135]取料块缩回位";
   IF #_w2 THEN "[324]取料块升降气缸" := TRUE; END_IF;
   #_w3 := #_w2 AND "[136]取料块下降位";
   IF #_w3 THEN
       "[327]取料块吸盘" := FALSE;
       "手动模式数据".S30放料块步骤 := 3.0;
   END_IF;
END_REGION

REGION Network 4: 复位
   RUNG wire#powerrail
      { S7_Templates := "SrcType := Real" } EQ_Contact(in1 := "手动模式数据".S30放料块步骤, in2 := 3.0)
      Contact( "[105]启动" )
      wire#w1
      R_Coil( "[324]取料块升降气缸" )
   END_RUNG
   RUNG wire#w1
      Contact( "[137]取料块上升位" )
      R_Coil( "[325]取料块伸缩气缸" )
   END_RUNG
   RUNG wire#w1
      Contact( "[137]取料块上升位" )
      Contact( "[135]取料块缩回位" )
      wire#w2
      Move(in := 0.0, out1 => "手动模式数据".S30放料块步骤)
   END_RUNG
   RUNG wire#w2
      Move(in := 3.0, out1 => "手动模式数据".手动总步骤)
   END_RUNG
   // the same network as SCL:
   #_w1 := ("手动模式数据".S30放料块步骤 = 3.0) AND "[105]启动";
   IF #_w1 THEN "[324]取料块升降气缸" := FALSE; END_IF;
   IF #_w1 AND "[137]取料块上升位" THEN "[325]取料块伸缩气缸" := FALSE; END_IF;
   IF #_w1 AND "[137]取料块上升位" AND "[135]取料块缩回位" THEN
       "手动模式数据".S30放料块步骤 := 0.0;
       "手动模式数据".手动总步骤 := 3.0;
   END_IF;
END_REGION
END_FUNCTION

FUNCTION "AI视觉信号映射" : Void   // FC21, LAD
{ S7_Optimized_Access := 'TRUE' }
VERSION : 0.1
BEGIN

REGION Network 1: Ai监视数据映射
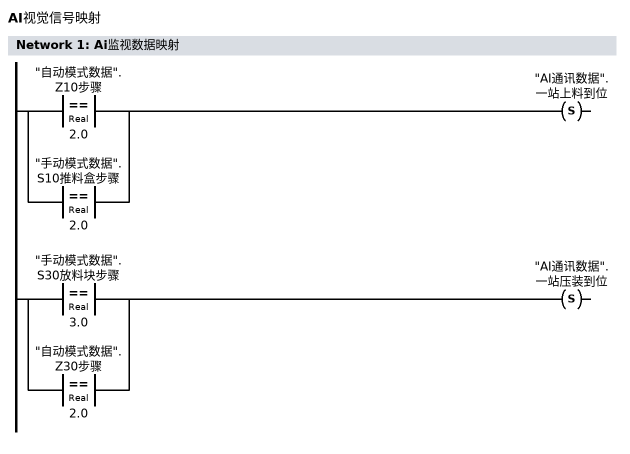
   RUNG wire#powerrail
      { S7_Templates := "SrcType := Real" } EQ_Contact(in1 := "自动模式数据".Z10步骤, in2 := 2.0)
      wire#w1
      S_Coil( "AI通讯数据".一站上料到位 )
   END_RUNG
   RUNG wire#powerrail
      { S7_Templates := "SrcType := Real" } EQ_Contact(in1 := "手动模式数据".S10推料盒步骤, in2 := 2.0)
   END_RUNG wire#w1
   RUNG wire#powerrail
      { S7_Templates := "SrcType := Real" } EQ_Contact(in1 := "手动模式数据".S30放料块步骤, in2 := 3.0)
      wire#w2
      S_Coil( "AI通讯数据".一站压装到位 )
   END_RUNG
   RUNG wire#powerrail
      { S7_Templates := "SrcType := Real" } EQ_Contact(in1 := "自动模式数据".Z30步骤, in2 := 2.0)
   END_RUNG wire#w2
   // the same network as SCL:
   IF ("自动模式数据".Z10步骤 = 2.0) OR ("手动模式数据".S10推料盒步骤 = 2.0) THEN "AI通讯数据".一站上料到位 := TRUE; END_IF;
   IF ("手动模式数据".S30放料块步骤 = 3.0) OR ("自动模式数据".Z30步骤 = 2.0) THEN "AI通讯数据".一站压装到位 := TRUE; END_IF;
END_REGION
END_FUNCTION

// folder: 自动模式

FUNCTION "Z10推料盒流程" : Void   // FC4, LAD
{ S7_Optimized_Access := 'TRUE' }
VERSION : 0.1
   VAR_TEMP   // added for the SCL form of the ladder/FBD networks
      _w1 : Bool;
      _w2 : Bool;
   END_VAR
BEGIN

REGION Network 1: 推出料盒
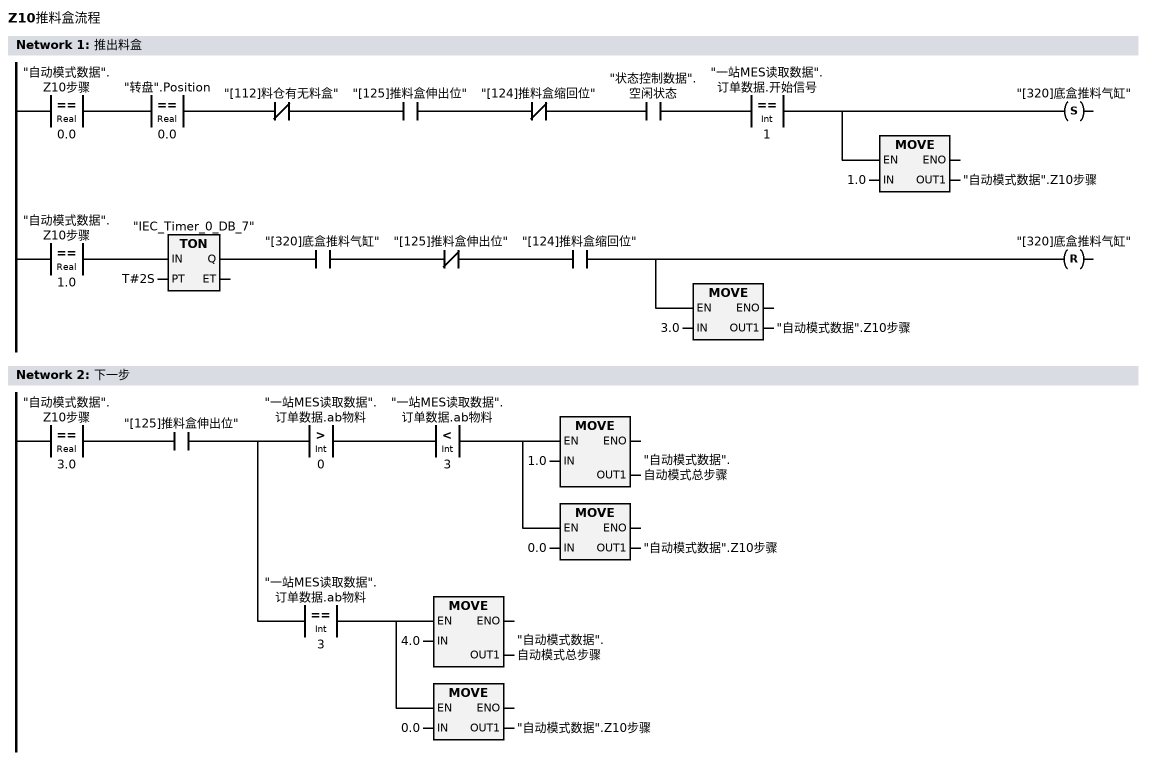
   #_w1 := ("自动模式数据".Z10步骤 = 0.0) AND ("转盘".Position = 0.0) AND NOT "[112]料仓有无料盒" AND "[125]推料盒伸出位" AND NOT "[124]推料盒缩回位" AND "状态控制数据".空闲状态 AND ("一站MES读取数据".订单数据.开始信号 = 1);
   IF #_w1 THEN
       "[320]底盒推料气缸" := TRUE;
       "自动模式数据".Z10步骤 := 1.0;
   END_IF;
   "IEC_Timer_0_DB_7".TON(IN := "自动模式数据".Z10步骤 = 1.0, PT := T#2S);
   #_w2 := "IEC_Timer_0_DB_7".Q AND "[320]底盒推料气缸" AND NOT "[125]推料盒伸出位" AND "[124]推料盒缩回位";
   IF #_w2 THEN
       "[320]底盒推料气缸" := FALSE;
       "自动模式数据".Z10步骤 := 3.0;
   END_IF;
END_REGION

REGION Network 2: 下一步
   RUNG wire#powerrail
      { S7_Templates := "SrcType := Real" } EQ_Contact(in1 := "自动模式数据".Z10步骤, in2 := 3.0)
      Contact( "[125]推料盒伸出位" )
      wire#w1
      { S7_Templates := "SrcType := Int" } GT_Contact(in1 := "一站MES读取数据".订单数据.ab物料, in2 := 0)
      { S7_Templates := "SrcType := Int" } LT_Contact(in1 := "一站MES读取数据".订单数据.ab物料, in2 := 3)
      wire#w2
      Move(in := 1.0, out1 => "自动模式数据".自动模式总步骤)
   END_RUNG
   RUNG wire#w2
      Move(in := 0.0, out1 => "自动模式数据".Z10步骤)
   END_RUNG
   RUNG wire#w1
      { S7_Templates := "SrcType := Int" } EQ_Contact(in1 := "一站MES读取数据".订单数据.ab物料, in2 := 3)
      wire#w3
      Move(in := 4.0, out1 => "自动模式数据".自动模式总步骤)
   END_RUNG
   RUNG wire#w3
      Move(in := 0.0, out1 => "自动模式数据".Z10步骤)
   END_RUNG
   // the same network as SCL:
   #_w1 := ("自动模式数据".Z10步骤 = 3.0) AND "[125]推料盒伸出位";
   IF #_w1 AND ("一站MES读取数据".订单数据.ab物料 > 0) AND ("一站MES读取数据".订单数据.ab物料 < 3) THEN
       "自动模式数据".自动模式总步骤 := 1.0;
       "自动模式数据".Z10步骤 := 0.0;
   END_IF;
   IF #_w1 AND ("一站MES读取数据".订单数据.ab物料 = 3) THEN
       "自动模式数据".自动模式总步骤 := 4.0;
       "自动模式数据".Z10步骤 := 0.0;
   END_IF;
END_REGION
END_FUNCTION

FUNCTION "Z20推料块流程" : Void   // FC11, LAD
{ S7_Optimized_Access := 'TRUE' }
VERSION : 0.1
   VAR_TEMP   // added for the SCL form of the ladder/FBD networks
      _w1 : Bool;
      _w2 : Bool;
      _w3 : Bool;
   END_VAR
BEGIN

REGION Network 1
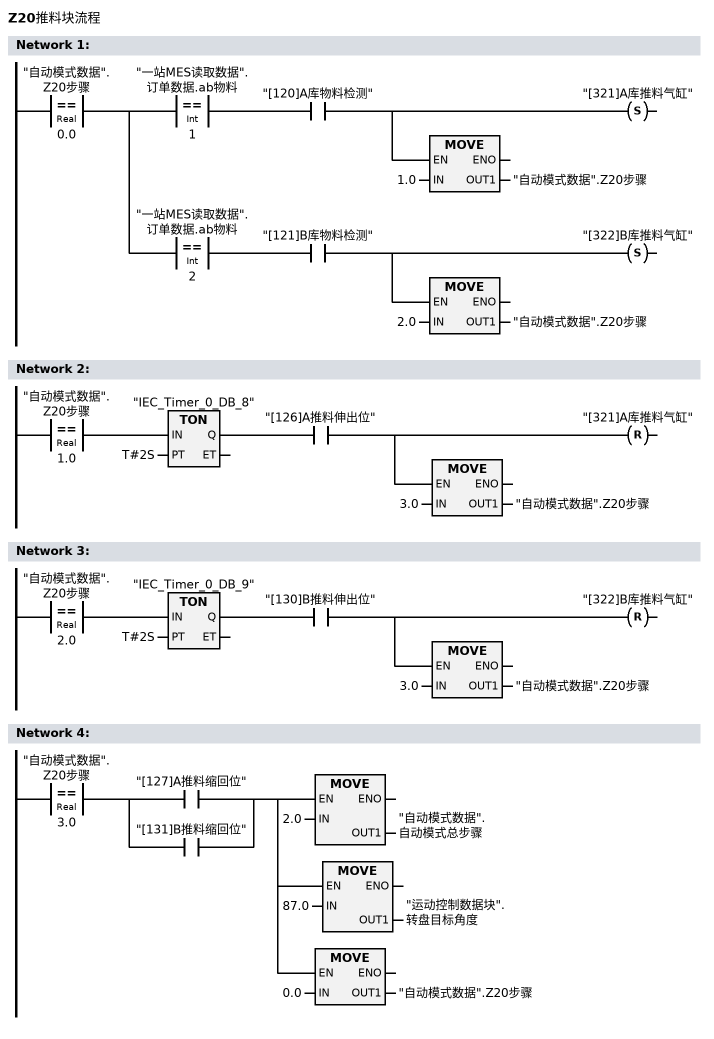
   RUNG wire#powerrail
      { S7_Templates := "SrcType := Real" } EQ_Contact(in1 := "自动模式数据".Z20步骤, in2 := 0.0)
      wire#w1
      { S7_Templates := "SrcType := Int" } EQ_Contact(in1 := "一站MES读取数据".订单数据.ab物料, in2 := 1)
      Contact( "[120]A库物料检测" )
      wire#w2
      S_Coil( "[321]A库推料气缸" )
   END_RUNG
   RUNG wire#w2
      Move(in := 1.0, out1 => "自动模式数据".Z20步骤)
   END_RUNG
   RUNG wire#w1
      { S7_Templates := "SrcType := Int" } EQ_Contact(in1 := "一站MES读取数据".订单数据.ab物料, in2 := 2)
      Contact( "[121]B库物料检测" )
      wire#w3
      S_Coil( "[322]B库推料气缸" )
   END_RUNG
   RUNG wire#w3
      Move(in := 2.0, out1 => "自动模式数据".Z20步骤)
   END_RUNG
   // the same network as SCL:
   #_w1 := "自动模式数据".Z20步骤 = 0.0;
   #_w2 := #_w1 AND ("一站MES读取数据".订单数据.ab物料 = 1) AND "[120]A库物料检测";
   IF #_w2 THEN
       "[321]A库推料气缸" := TRUE;
       "自动模式数据".Z20步骤 := 1.0;
   END_IF;
   #_w3 := #_w1 AND ("一站MES读取数据".订单数据.ab物料 = 2) AND "[121]B库物料检测";
   IF #_w3 THEN
       "[322]B库推料气缸" := TRUE;
       "自动模式数据".Z20步骤 := 2.0;
   END_IF;
END_REGION

REGION Network 2
   "IEC_Timer_0_DB_8".TON(IN := "自动模式数据".Z20步骤 = 1.0, PT := T#2S);
   #_w1 := "IEC_Timer_0_DB_8".Q AND "[126]A推料伸出位";
   IF #_w1 THEN
       "[321]A库推料气缸" := FALSE;
       "自动模式数据".Z20步骤 := 3.0;
   END_IF;
END_REGION

REGION Network 3
   "IEC_Timer_0_DB_9".TON(IN := "自动模式数据".Z20步骤 = 2.0, PT := T#2S);
   #_w1 := "IEC_Timer_0_DB_9".Q AND "[130]B推料伸出位";
   IF #_w1 THEN
       "[322]B库推料气缸" := FALSE;
       "自动模式数据".Z20步骤 := 3.0;
   END_IF;
END_REGION

REGION Network 4
   RUNG wire#powerrail
      { S7_Templates := "SrcType := Real" } EQ_Contact(in1 := "自动模式数据".Z20步骤, in2 := 3.0)
      wire#w1
      Contact( "[127]A推料缩回位" )
      wire#w2
      Move(in := 2.0, out1 => "自动模式数据".自动模式总步骤)
   END_RUNG
   RUNG wire#w1
      Contact( "[131]B推料缩回位" )
   END_RUNG wire#w2
   RUNG wire#w2
      Move(in := 87.0, out1 => "运动控制数据块".转盘目标角度)
   END_RUNG
   RUNG wire#w2
      Move(in := 0.0, out1 => "自动模式数据".Z20步骤)
   END_RUNG
   // the same network as SCL:
   IF ("自动模式数据".Z20步骤 = 3.0) AND ("[127]A推料缩回位" OR "[131]B推料缩回位") THEN
       "自动模式数据".自动模式总步骤 := 2.0;
       "运动控制数据块".转盘目标角度 := 87.0;
       "自动模式数据".Z20步骤 := 0.0;
   END_IF;
END_REGION
END_FUNCTION

FUNCTION "Z30取料块流程" : Void   // FC12, LAD
{ S7_Optimized_Access := 'TRUE' }
VERSION : 0.1
   VAR_TEMP   // added for the SCL form of the ladder/FBD networks
      _w1 : Bool;
      _w2 : Bool;
   END_VAR
BEGIN

REGION Network 1: 洗起来
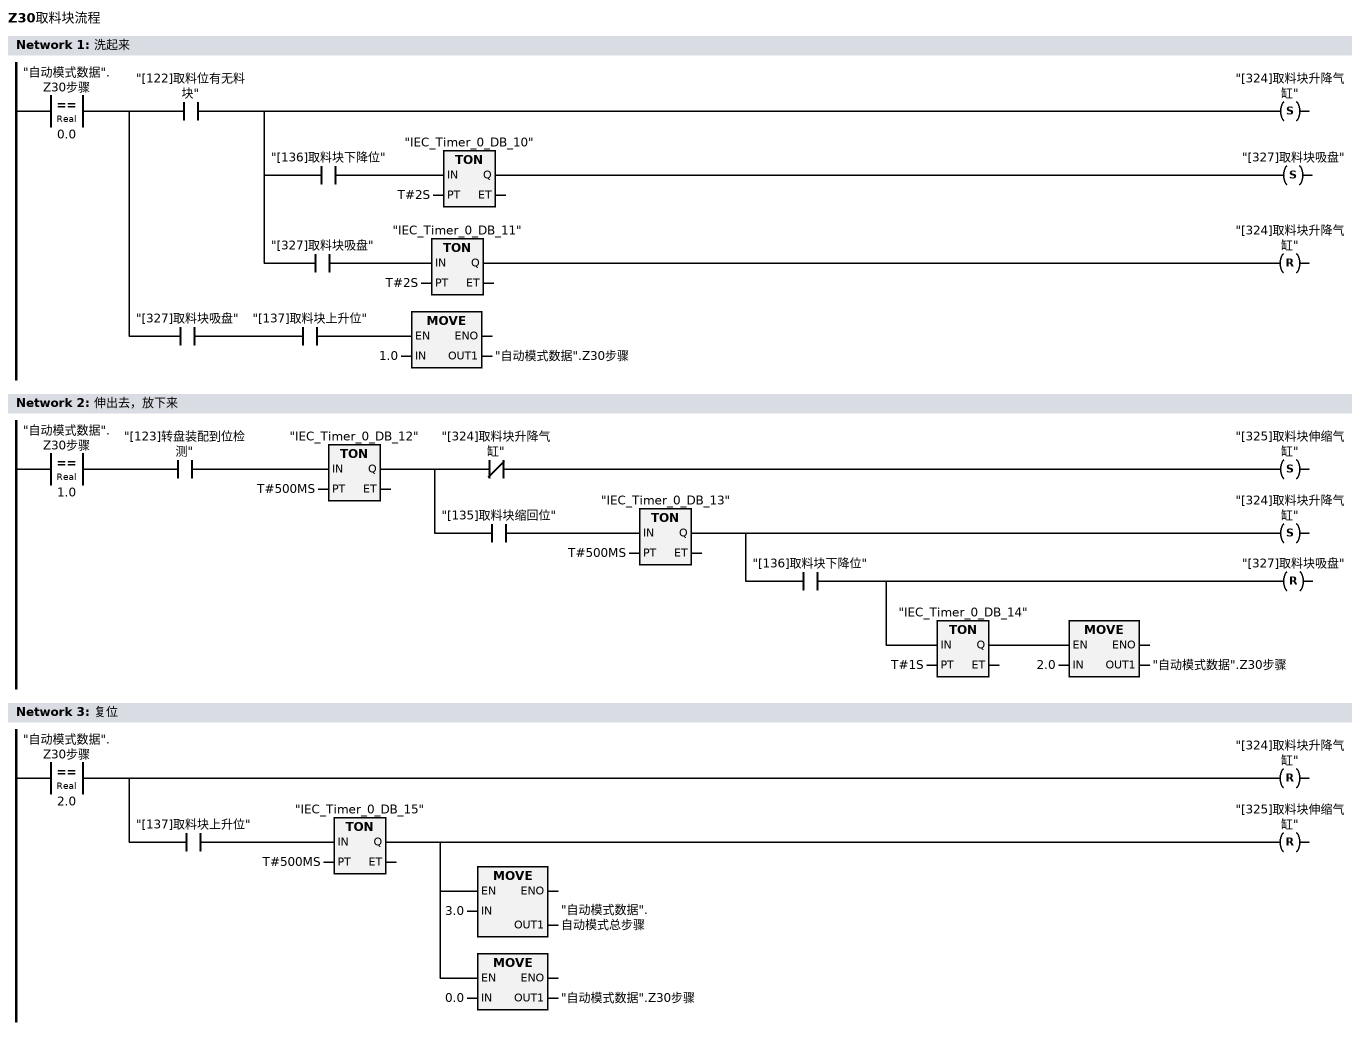
   #_w1 := "自动模式数据".Z30步骤 = 0.0;
   #_w2 := #_w1 AND "[122]取料位有无料块";
   IF #_w2 THEN "[324]取料块升降气缸" := TRUE; END_IF;
   "IEC_Timer_0_DB_10".TON(IN := #_w2 AND "[136]取料块下降位", PT := T#2S);
   IF "IEC_Timer_0_DB_10".Q THEN "[327]取料块吸盘" := TRUE; END_IF;
   "IEC_Timer_0_DB_11".TON(IN := #_w2 AND "[327]取料块吸盘", PT := T#2S);
   IF "IEC_Timer_0_DB_11".Q THEN "[324]取料块升降气缸" := FALSE; END_IF;
   IF #_w1 AND "[327]取料块吸盘" AND "[137]取料块上升位" THEN "自动模式数据".Z30步骤 := 1.0; END_IF;
END_REGION

REGION Network 2: 伸出去，放下来
   "IEC_Timer_0_DB_12".TON(IN := ("自动模式数据".Z30步骤 = 1.0) AND "[123]转盘装配到位检测", PT := T#500MS);
   IF "IEC_Timer_0_DB_12".Q AND NOT "[324]取料块升降气缸" THEN "[325]取料块伸缩气缸" := TRUE; END_IF;
   "IEC_Timer_0_DB_13".TON(IN := "IEC_Timer_0_DB_12".Q AND "[135]取料块缩回位", PT := T#500MS);
   IF "IEC_Timer_0_DB_13".Q THEN "[324]取料块升降气缸" := TRUE; END_IF;
   #_w1 := "IEC_Timer_0_DB_13".Q AND "[136]取料块下降位";
   IF #_w1 THEN "[327]取料块吸盘" := FALSE; END_IF;
   "IEC_Timer_0_DB_14".TON(IN := #_w1, PT := T#1S);
   IF "IEC_Timer_0_DB_14".Q THEN "自动模式数据".Z30步骤 := 2.0; END_IF;
END_REGION

REGION Network 3: 复位
   #_w1 := "自动模式数据".Z30步骤 = 2.0;
   IF #_w1 THEN "[324]取料块升降气缸" := FALSE; END_IF;
   "IEC_Timer_0_DB_15".TON(IN := #_w1 AND "[137]取料块上升位", PT := T#500MS);
   IF "IEC_Timer_0_DB_15".Q THEN
       "[325]取料块伸缩气缸" := FALSE;
       "自动模式数据".自动模式总步骤 := 3.0;
       "自动模式数据".Z30步骤 := 0.0;
   END_IF;
END_REGION
END_FUNCTION

FUNCTION "Z40A模式送料流程" : Void   // FC14, LAD
{ S7_Optimized_Access := 'TRUE' }
VERSION : 0.1
   VAR_TEMP   // added for the SCL form of the ladder/FBD networks
      _w1 : Bool;
      _w2 : Bool;
      _w3 : Bool;
   END_VAR
BEGIN

REGION Network 1
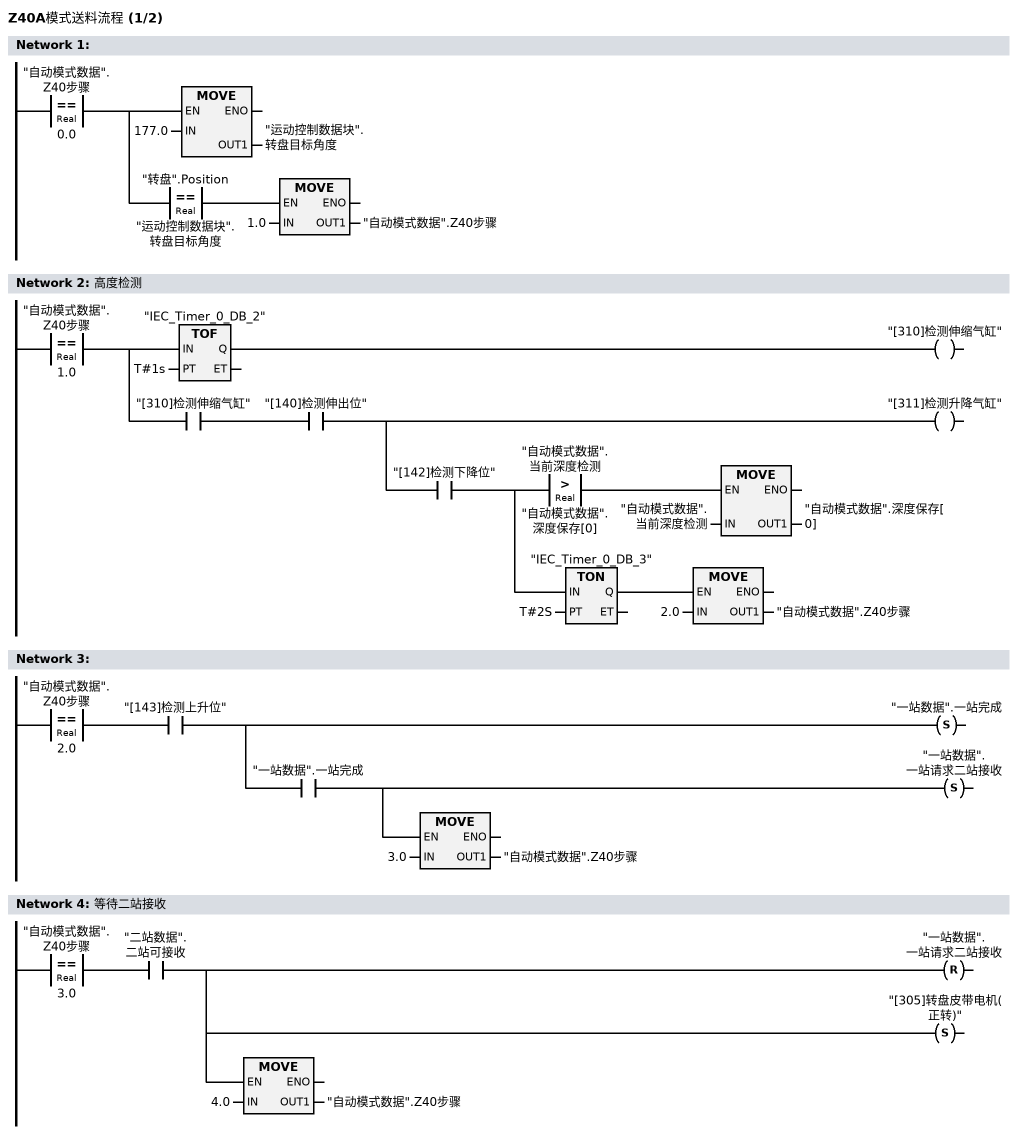
   RUNG wire#powerrail
      { S7_Templates := "SrcType := Real" } EQ_Contact(in1 := "自动模式数据".Z40步骤, in2 := 0.0)
      wire#w1
      Move(in := 177.0, out1 => "运动控制数据块".转盘目标角度)
   END_RUNG
   RUNG wire#w1
      { S7_Templates := "SrcType := Real" } EQ_Contact(in1 := "转盘".Position, in2 := "运动控制数据块".转盘目标角度)
      Move(in := 1.0, out1 => "自动模式数据".Z40步骤)
   END_RUNG
   // the same network as SCL:
   #_w1 := "自动模式数据".Z40步骤 = 0.0;
   IF #_w1 THEN "运动控制数据块".转盘目标角度 := 177.0; END_IF;
   IF #_w1 AND ("转盘".Position = "运动控制数据块".转盘目标角度) THEN "自动模式数据".Z40步骤 := 1.0; END_IF;
END_REGION

REGION Network 2: 高度检测
   #_w1 := "自动模式数据".Z40步骤 = 1.0;
   "IEC_Timer_0_DB_2".TOF(IN := #_w1, PT := T#1s);
   "[310]检测伸缩气缸" := "IEC_Timer_0_DB_2".Q;
   #_w2 := #_w1 AND "[310]检测伸缩气缸" AND "[140]检测伸出位";
   "[311]检测升降气缸" := #_w1 AND "[310]检测伸缩气缸" AND "[140]检测伸出位";
   #_w3 := #_w2 AND "[142]检测下降位";
   IF #_w3 AND ("自动模式数据".当前深度检测 > "自动模式数据".深度保存[0]) THEN "自动模式数据".深度保存[0] := "自动模式数据".当前深度检测; END_IF;
   "IEC_Timer_0_DB_3".TON(IN := #_w3, PT := T#2S);
   IF "IEC_Timer_0_DB_3".Q THEN "自动模式数据".Z40步骤 := 2.0; END_IF;
END_REGION

REGION Network 3
   RUNG wire#powerrail
      { S7_Templates := "SrcType := Real" } EQ_Contact(in1 := "自动模式数据".Z40步骤, in2 := 2.0)
      Contact( "[143]检测上升位" )
      wire#w1
      S_Coil( "一站数据".一站完成 )
   END_RUNG
   RUNG wire#w1
      Contact( "一站数据".一站完成 )
      wire#w2
      S_Coil( "一站数据".一站请求二站接收 )
   END_RUNG
   RUNG wire#w2
      Move(in := 3.0, out1 => "自动模式数据".Z40步骤)
   END_RUNG
   // the same network as SCL:
   #_w1 := ("自动模式数据".Z40步骤 = 2.0) AND "[143]检测上升位";
   IF #_w1 THEN "一站数据".一站完成 := TRUE; END_IF;
   IF #_w1 AND "一站数据".一站完成 THEN
       "一站数据".一站请求二站接收 := TRUE;
       "自动模式数据".Z40步骤 := 3.0;
   END_IF;
END_REGION

REGION Network 4: 等待二站接收
   RUNG wire#powerrail
      { S7_Templates := "SrcType := Real" } EQ_Contact(in1 := "自动模式数据".Z40步骤, in2 := 3.0)
      Contact( "二站数据".二站可接收 )
      wire#w1
      R_Coil( "一站数据".一站请求二站接收 )
   END_RUNG
   RUNG wire#w1
      S_Coil( "[305]转盘皮带电机(正转)" )
   END_RUNG
   RUNG wire#w1
      Move(in := 4.0, out1 => "自动模式数据".Z40步骤)
   END_RUNG
   // the same network as SCL:
   IF ("自动模式数据".Z40步骤 = 3.0) AND "二站数据".二站可接收 THEN
       "一站数据".一站请求二站接收 := FALSE;
       "[305]转盘皮带电机(正转)" := TRUE;
       "自动模式数据".Z40步骤 := 4.0;
   END_IF;
END_REGION

REGION Network 5
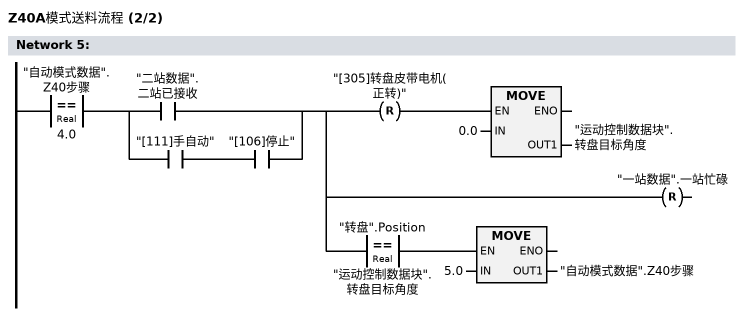
   RUNG wire#powerrail
      { S7_Templates := "SrcType := Real" } EQ_Contact(in1 := "自动模式数据".Z40步骤, in2 := 4.0)
      wire#w1
      Contact( "二站数据".二站已接收 )
      wire#w2
      R_Coil( "[305]转盘皮带电机(正转)" )
      Move(in := 0.0, out1 => "运动控制数据块".转盘目标角度)
   END_RUNG
   RUNG wire#w1
      Contact( "[111]手自动" )
      Contact( "[106]停止" )
   END_RUNG wire#w2
   RUNG wire#w2
      R_Coil( "一站数据".一站忙碌 )
   END_RUNG
   RUNG wire#w2
      { S7_Templates := "SrcType := Real" } EQ_Contact(in1 := "转盘".Position, in2 := "运动控制数据块".转盘目标角度)
      Move(in := 5.0, out1 => "自动模式数据".Z40步骤)
   END_RUNG
   // the same network as SCL:
   #_w1 := ("自动模式数据".Z40步骤 = 4.0) AND ("二站数据".二站已接收 OR ("[111]手自动" AND "[106]停止"));
   IF #_w1 THEN
       "[305]转盘皮带电机(正转)" := FALSE;
       "运动控制数据块".转盘目标角度 := 0.0;
       "一站数据".一站忙碌 := FALSE;
   END_IF;
   IF #_w1 AND ("转盘".Position = "运动控制数据块".转盘目标角度) THEN "自动模式数据".Z40步骤 := 5.0; END_IF;
END_REGION
END_FUNCTION

FUNCTION "Z50B模式送料流程" : Void   // FC15, LAD
{ S7_Optimized_Access := 'TRUE' }
VERSION : 0.1
// 不需要料块时，推出料盒后夹爪夹到第二站
   VAR_TEMP   // added for the SCL form of the ladder/FBD networks
      _w1 : Bool;
      _w2 : Bool;
   END_VAR
BEGIN

REGION Network 1: 到取料位
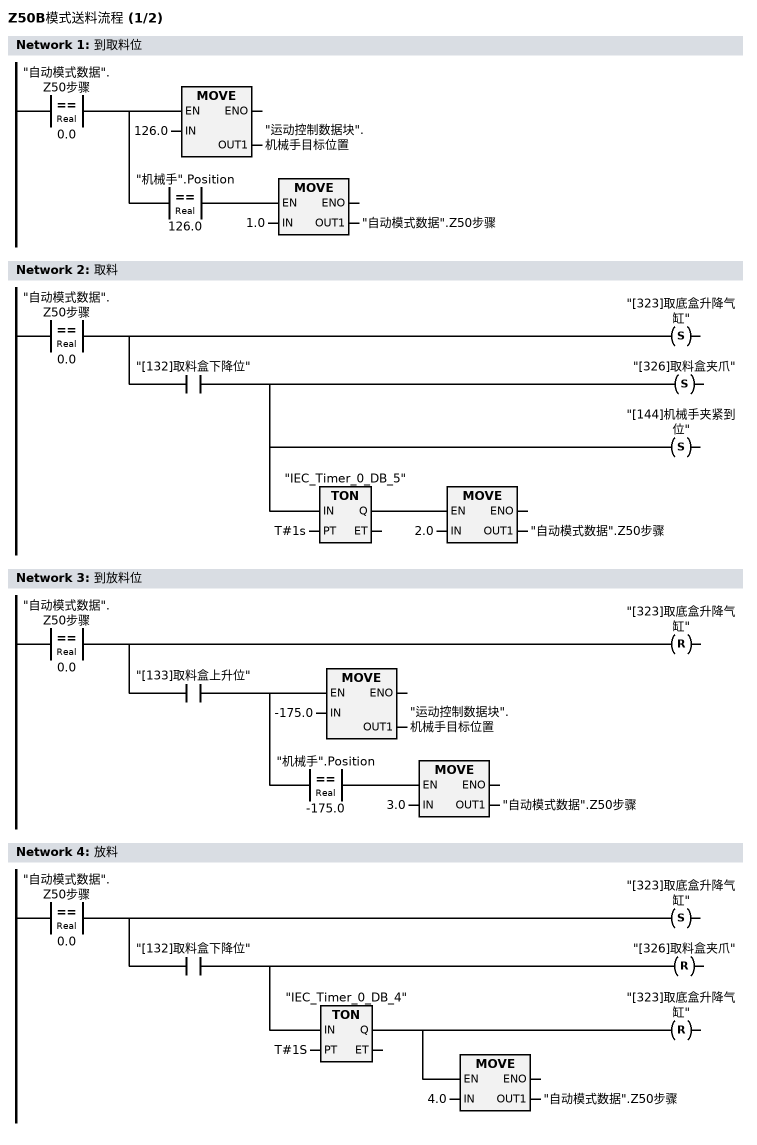
   RUNG wire#powerrail
      { S7_Templates := "SrcType := Real" } EQ_Contact(in1 := "自动模式数据".Z50步骤, in2 := 0.0)
      wire#w1
      Move(in := 126.0, out1 => "运动控制数据块".机械手目标位置)
   END_RUNG
   RUNG wire#w1
      { S7_Templates := "SrcType := Real" } EQ_Contact(in1 := "机械手".Position, in2 := 126.0)
      Move(in := 1.0, out1 => "自动模式数据".Z50步骤)
   END_RUNG
   // the same network as SCL:
   #_w1 := "自动模式数据".Z50步骤 = 0.0;
   IF #_w1 THEN "运动控制数据块".机械手目标位置 := 126.0; END_IF;
   IF #_w1 AND ("机械手".Position = 126.0) THEN "自动模式数据".Z50步骤 := 1.0; END_IF;
END_REGION

REGION Network 2: 取料
   #_w1 := "自动模式数据".Z50步骤 = 0.0;
   IF #_w1 THEN "[323]取底盒升降气缸" := TRUE; END_IF;
   #_w2 := #_w1 AND "[132]取料盒下降位";
   IF #_w2 THEN
       "[326]取料盒夹爪" := TRUE;
       "[144]机械手夹紧到位" := TRUE;
   END_IF;
   "IEC_Timer_0_DB_5".TON(IN := #_w2, PT := T#1s);
   IF "IEC_Timer_0_DB_5".Q THEN "自动模式数据".Z50步骤 := 2.0; END_IF;
END_REGION

REGION Network 3: 到放料位
   RUNG wire#powerrail
      { S7_Templates := "SrcType := Real" } EQ_Contact(in1 := "自动模式数据".Z50步骤, in2 := 0.0)
      wire#w1
      R_Coil( "[323]取底盒升降气缸" )
   END_RUNG
   RUNG wire#w1
      Contact( "[133]取料盒上升位" )
      wire#w2
      Move(in := -175.0, out1 => "运动控制数据块".机械手目标位置)
   END_RUNG
   RUNG wire#w2
      { S7_Templates := "SrcType := Real" } EQ_Contact(in1 := "机械手".Position, in2 := -175.0)
      Move(in := 3.0, out1 => "自动模式数据".Z50步骤)
   END_RUNG
   // the same network as SCL:
   #_w1 := "自动模式数据".Z50步骤 = 0.0;
   IF #_w1 THEN "[323]取底盒升降气缸" := FALSE; END_IF;
   #_w2 := #_w1 AND "[133]取料盒上升位";
   IF #_w2 THEN "运动控制数据块".机械手目标位置 := -175.0; END_IF;
   IF #_w2 AND ("机械手".Position = (-175.0)) THEN "自动模式数据".Z50步骤 := 3.0; END_IF;
END_REGION

REGION Network 4: 放料
   #_w1 := "自动模式数据".Z50步骤 = 0.0;
   IF #_w1 THEN "[323]取底盒升降气缸" := TRUE; END_IF;
   #_w2 := #_w1 AND "[132]取料盒下降位";
   IF #_w2 THEN "[326]取料盒夹爪" := FALSE; END_IF;
   "IEC_Timer_0_DB_4".TON(IN := #_w2, PT := T#1S);
   IF "IEC_Timer_0_DB_4".Q THEN
       "[323]取底盒升降气缸" := FALSE;
       "自动模式数据".Z50步骤 := 4.0;
   END_IF;
END_REGION

REGION Network 5: 复位
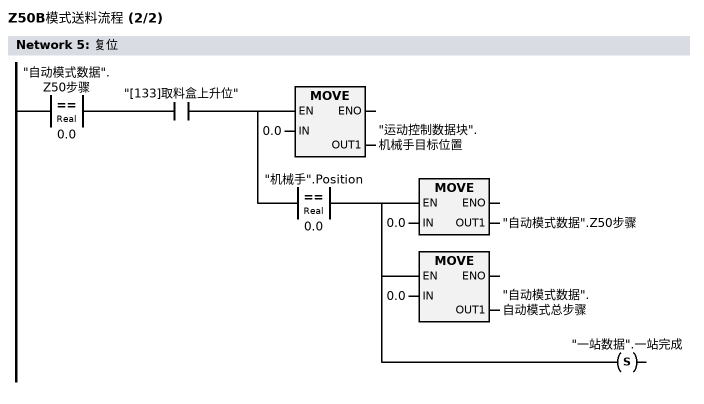
   RUNG wire#powerrail
      { S7_Templates := "SrcType := Real" } EQ_Contact(in1 := "自动模式数据".Z50步骤, in2 := 0.0)
      Contact( "[133]取料盒上升位" )
      wire#w1
      Move(in := 0.0, out1 => "运动控制数据块".机械手目标位置)
   END_RUNG
   RUNG wire#w1
      { S7_Templates := "SrcType := Real" } EQ_Contact(in1 := "机械手".Position, in2 := 0.0)
      wire#w2
      Move(in := 0.0, out1 => "自动模式数据".Z50步骤)
   END_RUNG
   RUNG wire#w2
      Move(in := 0.0, out1 => "自动模式数据".自动模式总步骤)
   END_RUNG
   RUNG wire#w2
      S_Coil( "一站数据".一站完成 )
   END_RUNG
   // the same network as SCL:
   #_w1 := ("自动模式数据".Z50步骤 = 0.0) AND "[133]取料盒上升位";
   IF #_w1 THEN "运动控制数据块".机械手目标位置 := 0.0; END_IF;
   IF #_w1 AND ("机械手".Position = 0.0) THEN
       "自动模式数据".Z50步骤 := 0.0;
       "自动模式数据".自动模式总步骤 := 0.0;
       "一站数据".一站完成 := TRUE;
   END_IF;
END_REGION
END_FUNCTION

FUNCTION "数据转换以及检测" : Void   // FC17, LAD
{ S7_Optimized_Access := 'TRUE' }
VERSION : 0.1
   VAR_TEMP   // added for the SCL form of the ladder/FBD networks
      _w1 : Bool;
      _w2 : Bool;
      _w3 : Bool;
   END_VAR
BEGIN

REGION Network 1: 原始数据转换
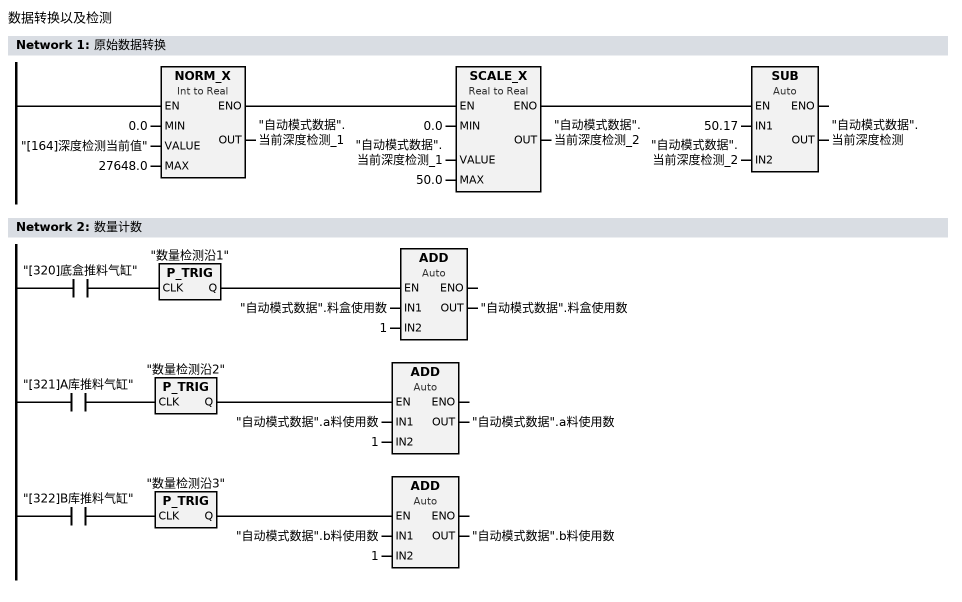
   RUNG wire#powerrail
      { S7_Templates := "[SrcType := Int, DestType := Real]" } Normalize(min := 0.0, value := "[164]深度检测当前值", max := 27648.0, out => "自动模式数据".当前深度检测_1)
      { S7_Templates := "[SrcType := Real, DestType := Real]" } Scale(min := 0.0, value := "自动模式数据".当前深度检测_1, max := 50.0, out => "自动模式数据".当前深度检测_2)
      Sub(in1 := 50.17, in2 := "自动模式数据".当前深度检测_2, out => "自动模式数据".当前深度检测)
   END_RUNG
   // the same network as SCL:
   "自动模式数据".当前深度检测_1 := NORM_X(MIN := 0.0, VALUE := "[164]深度检测当前值", MAX := 27648.0);
   "自动模式数据".当前深度检测_2 := SCALE_X(MIN := 0.0, VALUE := "自动模式数据".当前深度检测_1, MAX := 50.0);
   "自动模式数据".当前深度检测 := 50.17 - "自动模式数据".当前深度检测_2;
END_REGION

REGION Network 2: 数量计数
   RUNG wire#powerrail
      Contact( "[320]底盒推料气缸" )
      P_Trig( "数量检测沿1" )
      Add(in1 := "自动模式数据".料盒使用数, in2 := 1, out => "自动模式数据".料盒使用数)
   END_RUNG
   RUNG wire#powerrail
      Contact( "[321]A库推料气缸" )
      P_Trig( "数量检测沿2" )
      Add(in1 := "自动模式数据".a料使用数, in2 := 1, out => "自动模式数据".a料使用数)
   END_RUNG
   RUNG wire#powerrail
      Contact( "[322]B库推料气缸" )
      P_Trig( "数量检测沿3" )
      Add(in1 := "自动模式数据".b料使用数, in2 := 1, out => "自动模式数据".b料使用数)
   END_RUNG
   // the same network as SCL:
   #_w1 := "[320]底盒推料气缸" AND NOT "数量检测沿1";   // rising edge
   "数量检测沿1" := "[320]底盒推料气缸";
   IF #_w1 THEN "自动模式数据".料盒使用数 := "自动模式数据".料盒使用数 + 1; END_IF;
   #_w2 := "[321]A库推料气缸" AND NOT "数量检测沿2";   // rising edge
   "数量检测沿2" := "[321]A库推料气缸";
   IF #_w2 THEN "自动模式数据".a料使用数 := "自动模式数据".a料使用数 + 1; END_IF;
   #_w3 := "[322]B库推料气缸" AND NOT "数量检测沿3";   // rising edge
   "数量检测沿3" := "[322]B库推料气缸";
   IF #_w3 THEN "自动模式数据".b料使用数 := "自动模式数据".b料使用数 + 1; END_IF;
END_REGION
END_FUNCTION

// folder: 运动控制

FUNCTION "转盘程序" : Void   // FC1, LAD
{ S7_Optimized_Access := 'TRUE' }
VERSION : 0.1
BEGIN

REGION Network 1
